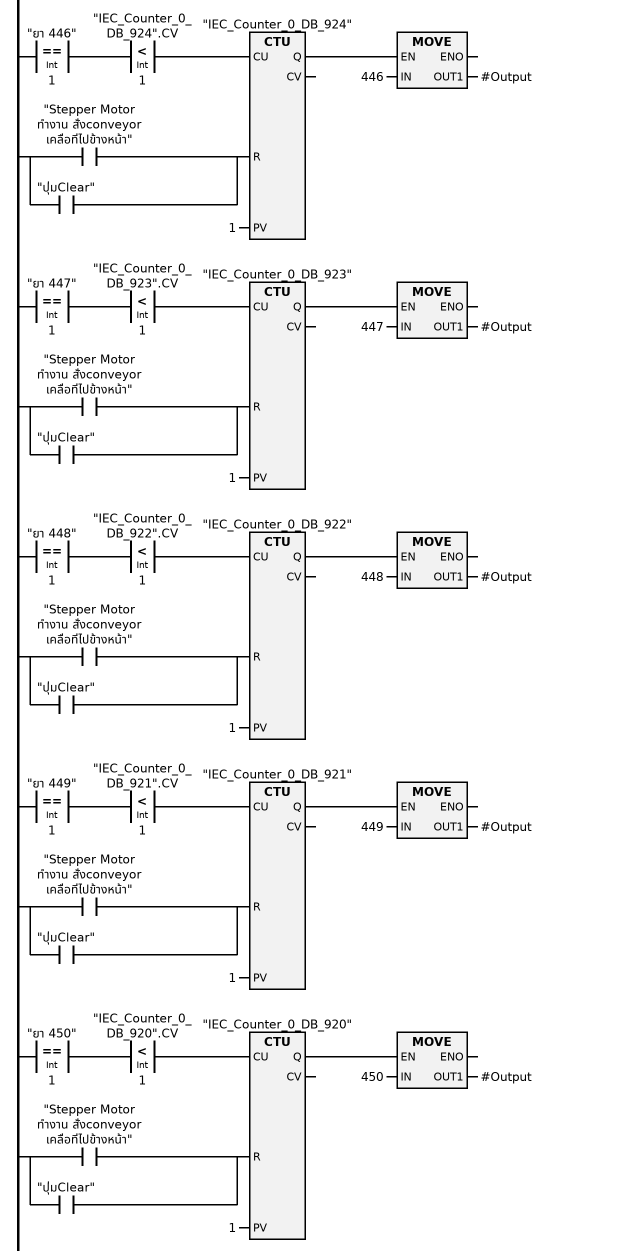
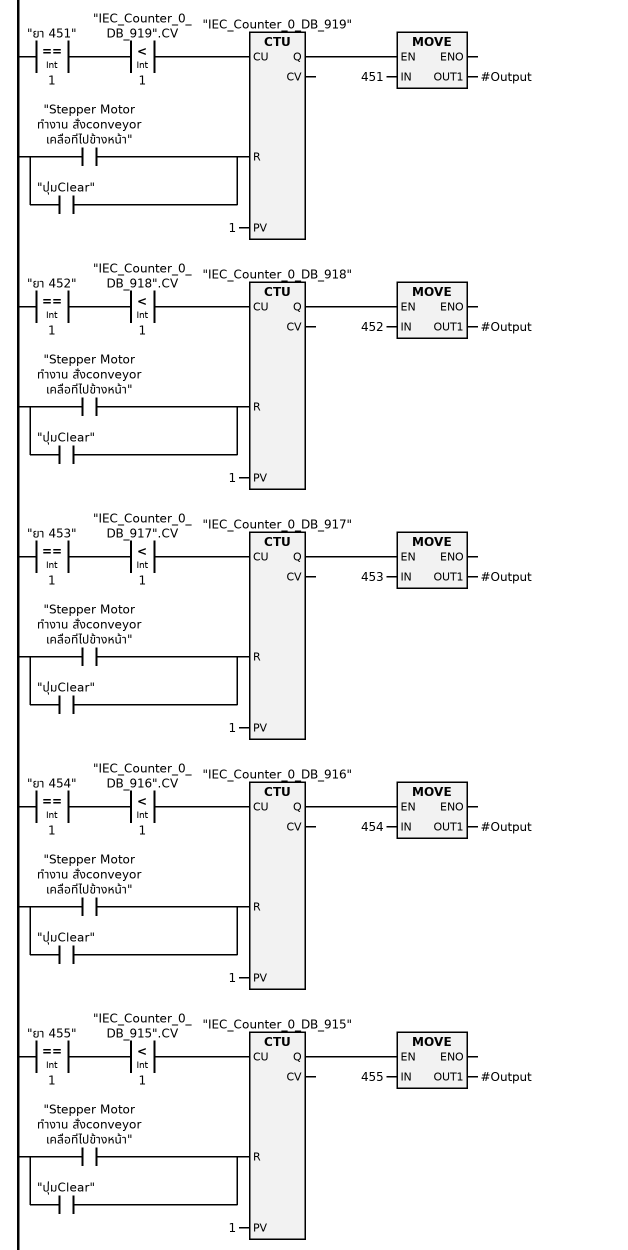
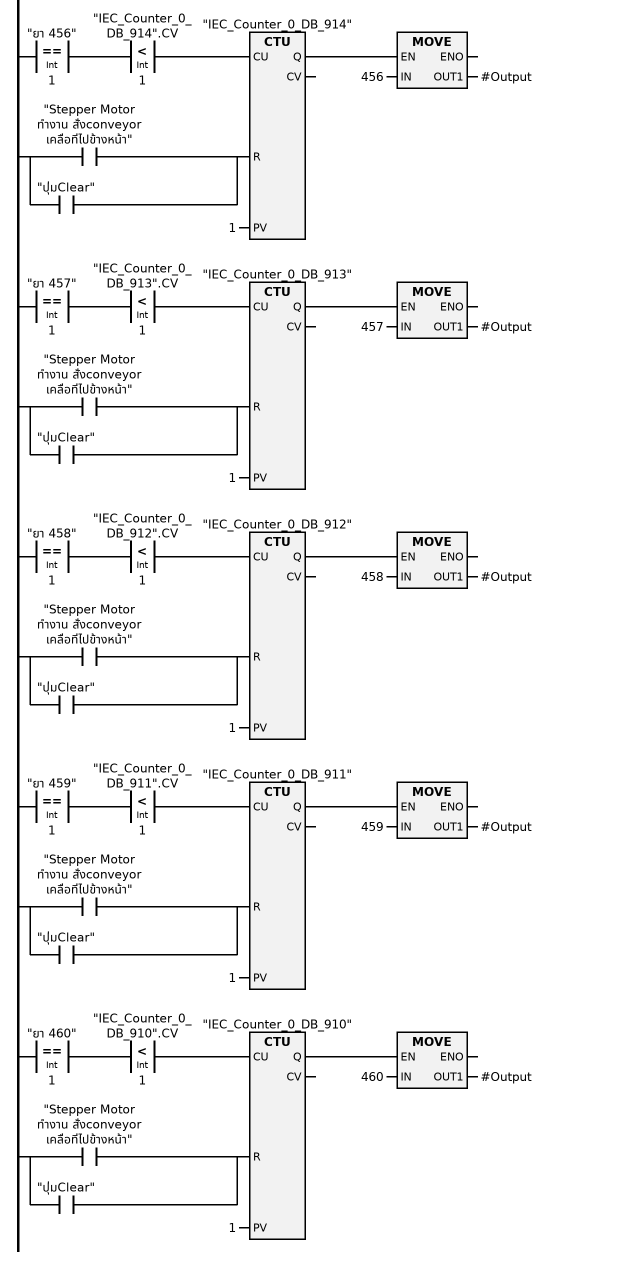
   "IEC_Counter_0_DB_929".CTU(CU := ("ยา 441" = 1) AND ("IEC_Counter_0_DB_929".CV < 1),
                           R := "Stepper Motor ทำงาน สั่งconveyor เคลื่อที่ไปข้างหน้า" OR "ปุ่มClear",
                           PV := 1);
   IF "IEC_Counter_0_DB_929".Q THEN #Output := 441; END_IF;
   "IEC_Counter_0_DB_928".CTU(CU := ("ยา 442" = 1) AND ("IEC_Counter_0_DB_928".CV < 1),
                           R := "Stepper Motor ทำงาน สั่งconveyor เคลื่อที่ไปข้างหน้า" OR "ปุ่มClear",
                           PV := 1);
   IF "IEC_Counter_0_DB_928".Q THEN #Output := 442; END_IF;
   "IEC_Counter_0_DB_927".CTU(CU := ("ยา 443" = 1) AND ("IEC_Counter_0_DB_927".CV < 1),
                           R := "Stepper Motor ทำงาน สั่งconveyor เคลื่อที่ไปข้างหน้า" OR "ปุ่มClear",
                           PV := 1);
   IF "IEC_Counter_0_DB_927".Q THEN #Output := 443; END_IF;
   "IEC_Counter_0_DB_926".CTU(CU := ("ยา 444" = 1) AND ("IEC_Counter_0_DB_926".CV < 1),
                           R := "Stepper Motor ทำงาน สั่งconveyor เคลื่อที่ไปข้างหน้า" OR "ปุ่มClear",
                           PV := 1);
   IF "IEC_Counter_0_DB_926".Q THEN #Output := 444; END_IF;
   "IEC_Counter_0_DB_925".CTU(CU := ("ยา 445" = 1) AND ("IEC_Counter_0_DB_925".CV < 1),
                           R := "Stepper Motor ทำงาน สั่งconveyor เคลื่อที่ไปข้างหน้า" OR "ปุ่มClear",
                           PV := 1);
   IF "IEC_Counter_0_DB_925".Q THEN #Output := 445; END_IF;
   "IEC_Counter_0_DB_924".CTU(CU := ("ยา 446" = 1) AND ("IEC_Counter_0_DB_924".CV < 1),
                           R := "Stepper Motor ทำงาน สั่งconveyor เคลื่อที่ไปข้างหน้า" OR "ปุ่มClear",
                           PV := 1);
   IF "IEC_Counter_0_DB_924".Q THEN #Output := 446; END_IF;
   "IEC_Counter_0_DB_923".CTU(CU := ("ยา 447" = 1) AND ("IEC_Counter_0_DB_923".CV < 1),
                           R := "Stepper Motor ทำงาน สั่งconveyor เคลื่อที่ไปข้างหน้า" OR "ปุ่มClear",
                           PV := 1);
   IF "IEC_Counter_0_DB_923".Q THEN #Output := 447; END_IF;
   "IEC_Counter_0_DB_922".CTU(CU := ("ยา 448" = 1) AND ("IEC_Counter_0_DB_922".CV < 1),
                           R := "Stepper Motor ทำงาน สั่งconveyor เคลื่อที่ไปข้างหน้า" OR "ปุ่มClear",
                           PV := 1);
   IF "IEC_Counter_0_DB_922".Q THEN #Output := 448; END_IF;
   "IEC_Counter_0_DB_921".CTU(CU := ("ยา 449" = 1) AND ("IEC_Counter_0_DB_921".CV < 1),
                           R := "Stepper Motor ทำงาน สั่งconveyor เคลื่อที่ไปข้างหน้า" OR "ปุ่มClear",
                           PV := 1);
   IF "IEC_Counter_0_DB_921".Q THEN #Output := 449; END_IF;
   "IEC_Counter_0_DB_920".CTU(CU := ("ยา 450" = 1) AND ("IEC_Counter_0_DB_920".CV < 1),
                           R := "Stepper Motor ทำงาน สั่งconveyor เคลื่อที่ไปข้างหน้า" OR "ปุ่มClear",
                           PV := 1);
   IF "IEC_Counter_0_DB_920".Q THEN #Output := 450; END_IF;
   "IEC_Counter_0_DB_919".CTU(CU := ("ยา 451" = 1) AND ("IEC_Counter_0_DB_919".CV < 1),
                           R := "Stepper Motor ทำงาน สั่งconveyor เคลื่อที่ไปข้างหน้า" OR "ปุ่มClear",
                           PV := 1);
   IF "IEC_Counter_0_DB_919".Q THEN #Output := 451; END_IF;
   "IEC_Counter_0_DB_918".CTU(CU := ("ยา 452" = 1) AND ("IEC_Counter_0_DB_918".CV < 1),
                           R := "Stepper Motor ทำงาน สั่งconveyor เคลื่อที่ไปข้างหน้า" OR "ปุ่มClear",
                           PV := 1);
   IF "IEC_Counter_0_DB_918".Q THEN #Output := 452; END_IF;
   "IEC_Counter_0_DB_917".CTU(CU := ("ยา 453" = 1) AND ("IEC_Counter_0_DB_917".CV < 1),
                           R := "Stepper Motor ทำงาน สั่งconveyor เคลื่อที่ไปข้างหน้า" OR "ปุ่มClear",
                           PV := 1);
   IF "IEC_Counter_0_DB_917".Q THEN #Output := 453; END_IF;
   "IEC_Counter_0_DB_916".CTU(CU := ("ยา 454" = 1) AND ("IEC_Counter_0_DB_916".CV < 1),
                           R := "Stepper Motor ทำงาน สั่งconveyor เคลื่อที่ไปข้างหน้า" OR "ปุ่มClear",
                           PV := 1);
   IF "IEC_Counter_0_DB_916".Q THEN #Output := 454; END_IF;
   "IEC_Counter_0_DB_915".CTU(CU := ("ยา 455" = 1) AND ("IEC_Counter_0_DB_915".CV < 1),
                           R := "Stepper Motor ทำงาน สั่งconveyor เคลื่อที่ไปข้างหน้า" OR "ปุ่มClear",
                           PV := 1);
   IF "IEC_Counter_0_DB_915".Q THEN #Output := 455; END_IF;
   "IEC_Counter_0_DB_914".CTU(CU := ("ยา 456" = 1) AND ("IEC_Counter_0_DB_914".CV < 1),
                           R := "Stepper Motor ทำงาน สั่งconveyor เคลื่อที่ไปข้างหน้า" OR "ปุ่มClear",
                           PV := 1);
   IF "IEC_Counter_0_DB_914".Q THEN #Output := 456; END_IF;
   "IEC_Counter_0_DB_913".CTU(CU := ("ยา 457" = 1) AND ("IEC_Counter_0_DB_913".CV < 1),
                           R := "Stepper Motor ทำงาน สั่งconveyor เคลื่อที่ไปข้างหน้า" OR "ปุ่มClear",
                           PV := 1);
   IF "IEC_Counter_0_DB_913".Q THEN #Output := 457; END_IF;
   "IEC_Counter_0_DB_912".CTU(CU := ("ยา 458" = 1) AND ("IEC_Counter_0_DB_912".CV < 1),
                           R := "Stepper Motor ทำงาน สั่งconveyor เคลื่อที่ไปข้างหน้า" OR "ปุ่มClear",
                           PV := 1);
   IF "IEC_Counter_0_DB_912".Q THEN #Output := 458; END_IF;
   "IEC_Counter_0_DB_911".CTU(CU := ("ยา 459" = 1) AND ("IEC_Counter_0_DB_911".CV < 1),
                           R := "Stepper Motor ทำงาน สั่งconveyor เคลื่อที่ไปข้างหน้า" OR "ปุ่มClear",
                           PV := 1);
   IF "IEC_Counter_0_DB_911".Q THEN #Output := 459; END_IF;
   "IEC_Counter_0_DB_910".CTU(CU := ("ยา 460" = 1) AND ("IEC_Counter_0_DB_910".CV < 1),
                           R := "Stepper Motor ทำงาน สั่งconveyor เคลื่อที่ไปข้างหน้า" OR "ปุ่มClear",
                           PV := 1);
   IF "IEC_Counter_0_DB_910".Q THEN #Output := 460; END_IF;
END_REGION

REGION Network 24
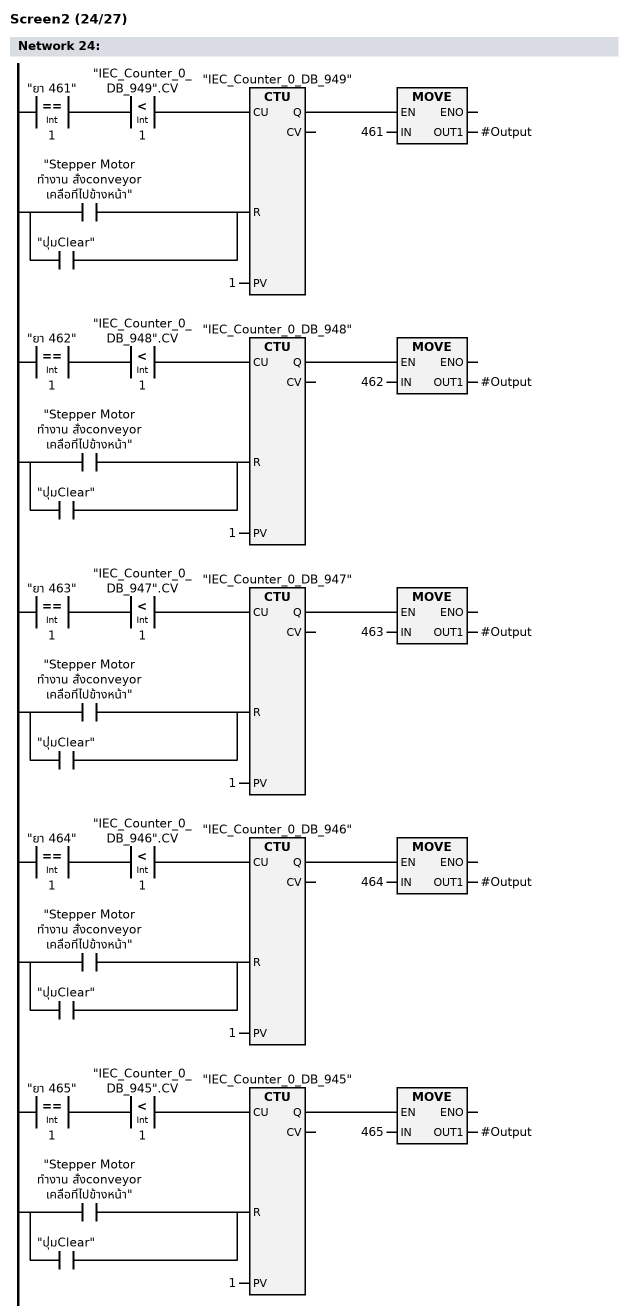
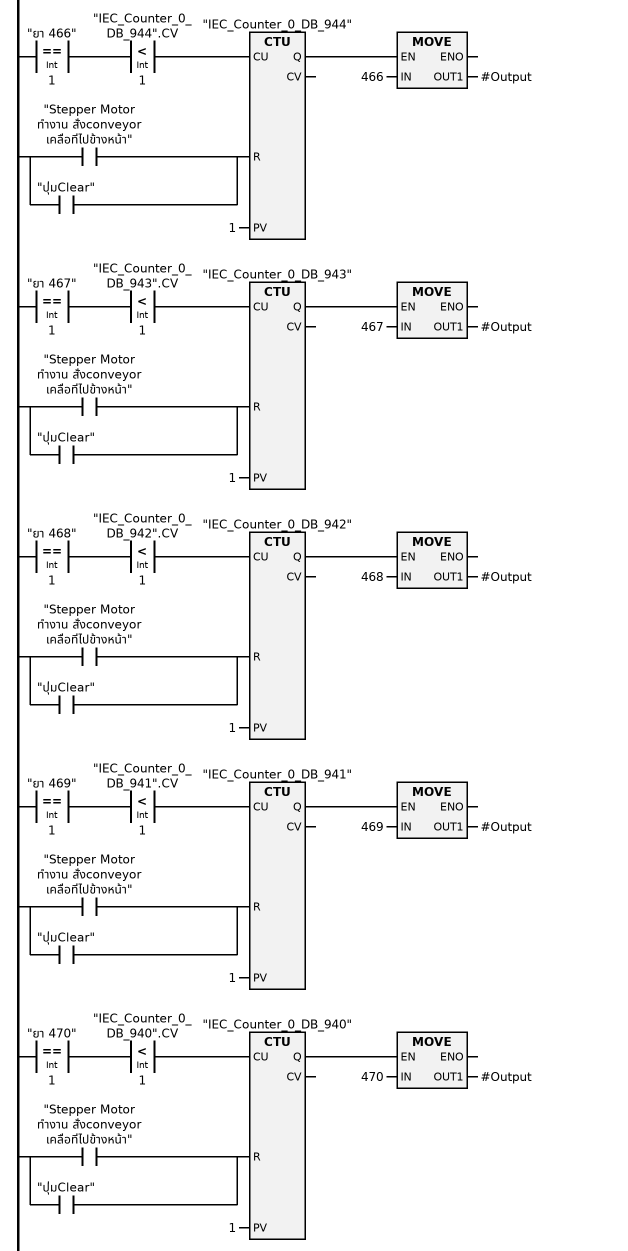
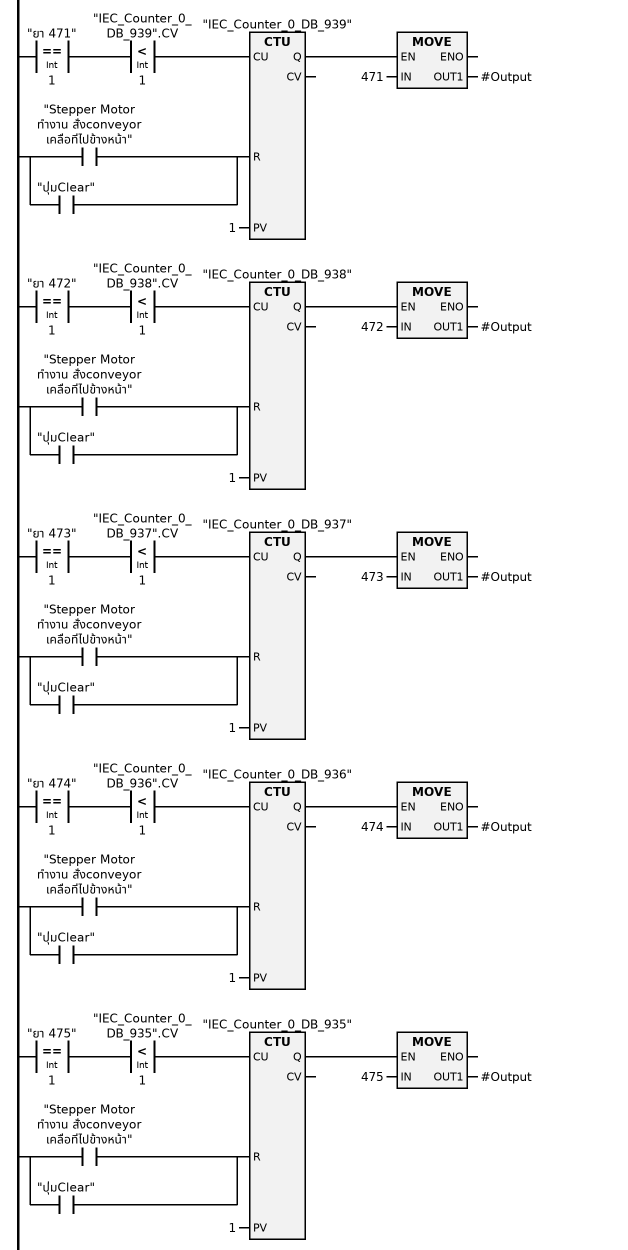
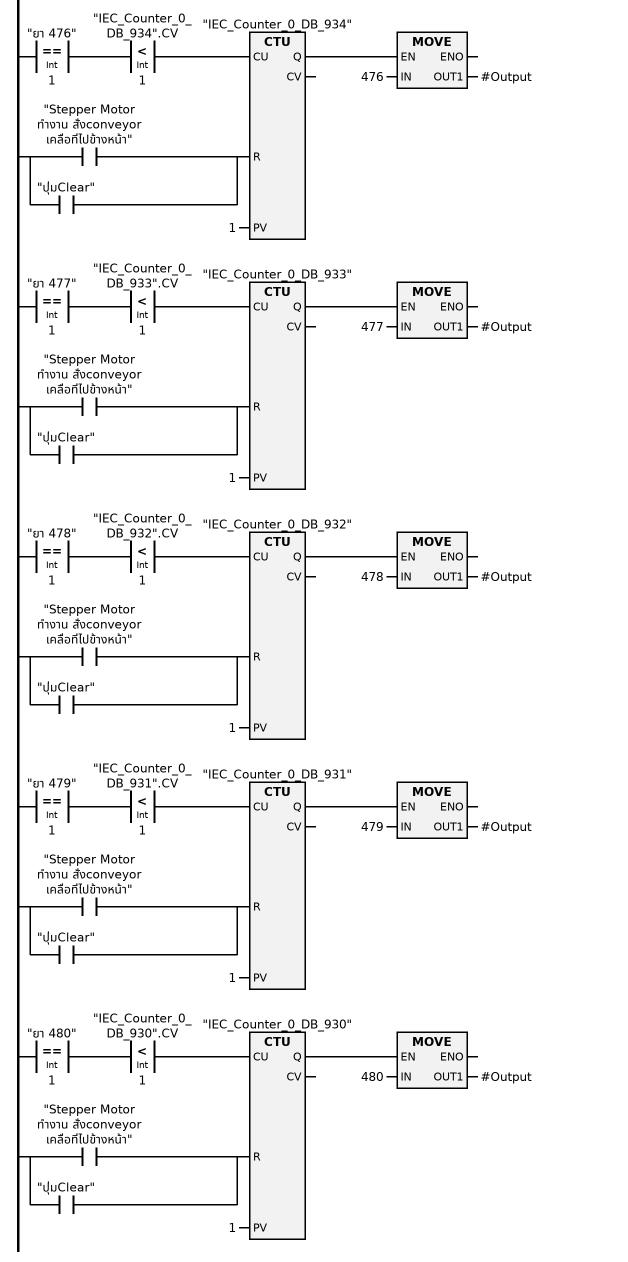
   "IEC_Counter_0_DB_949".CTU(CU := ("ยา 461" = 1) AND ("IEC_Counter_0_DB_949".CV < 1),
                           R := "Stepper Motor ทำงาน สั่งconveyor เคลื่อที่ไปข้างหน้า" OR "ปุ่มClear",
                           PV := 1);
   IF "IEC_Counter_0_DB_949".Q THEN #Output := 461; END_IF;
   "IEC_Counter_0_DB_948".CTU(CU := ("ยา 462" = 1) AND ("IEC_Counter_0_DB_948".CV < 1),
                           R := "Stepper Motor ทำงาน สั่งconveyor เคลื่อที่ไปข้างหน้า" OR "ปุ่มClear",
                           PV := 1);
   IF "IEC_Counter_0_DB_948".Q THEN #Output := 462; END_IF;
   "IEC_Counter_0_DB_947".CTU(CU := ("ยา 463" = 1) AND ("IEC_Counter_0_DB_947".CV < 1),
                           R := "Stepper Motor ทำงาน สั่งconveyor เคลื่อที่ไปข้างหน้า" OR "ปุ่มClear",
                           PV := 1);
   IF "IEC_Counter_0_DB_947".Q THEN #Output := 463; END_IF;
   "IEC_Counter_0_DB_946".CTU(CU := ("ยา 464" = 1) AND ("IEC_Counter_0_DB_946".CV < 1),
                           R := "Stepper Motor ทำงาน สั่งconveyor เคลื่อที่ไปข้างหน้า" OR "ปุ่มClear",
                           PV := 1);
   IF "IEC_Counter_0_DB_946".Q THEN #Output := 464; END_IF;
   "IEC_Counter_0_DB_945".CTU(CU := ("ยา 465" = 1) AND ("IEC_Counter_0_DB_945".CV < 1),
                           R := "Stepper Motor ทำงาน สั่งconveyor เคลื่อที่ไปข้างหน้า" OR "ปุ่มClear",
                           PV := 1);
   IF "IEC_Counter_0_DB_945".Q THEN #Output := 465; END_IF;
   "IEC_Counter_0_DB_944".CTU(CU := ("ยา 466" = 1) AND ("IEC_Counter_0_DB_944".CV < 1),
                           R := "Stepper Motor ทำงาน สั่งconveyor เคลื่อที่ไปข้างหน้า" OR "ปุ่มClear",
                           PV := 1);
   IF "IEC_Counter_0_DB_944".Q THEN #Output := 466; END_IF;
   "IEC_Counter_0_DB_943".CTU(CU := ("ยา 467" = 1) AND ("IEC_Counter_0_DB_943".CV < 1),
                           R := "Stepper Motor ทำงาน สั่งconveyor เคลื่อที่ไปข้างหน้า" OR "ปุ่มClear",
                           PV := 1);
   IF "IEC_Counter_0_DB_943".Q THEN #Output := 467; END_IF;
   "IEC_Counter_0_DB_942".CTU(CU := ("ยา 468" = 1) AND ("IEC_Counter_0_DB_942".CV < 1),
                           R := "Stepper Motor ทำงาน สั่งconveyor เคลื่อที่ไปข้างหน้า" OR "ปุ่มClear",
                           PV := 1);
   IF "IEC_Counter_0_DB_942".Q THEN #Output := 468; END_IF;
   "IEC_Counter_0_DB_941".CTU(CU := ("ยา 469" = 1) AND ("IEC_Counter_0_DB_941".CV < 1),
                           R := "Stepper Motor ทำงาน สั่งconveyor เคลื่อที่ไปข้างหน้า" OR "ปุ่มClear",
                           PV := 1);
   IF "IEC_Counter_0_DB_941".Q THEN #Output := 469; END_IF;
   "IEC_Counter_0_DB_940".CTU(CU := ("ยา 470" = 1) AND ("IEC_Counter_0_DB_940".CV < 1),
                           R := "Stepper Motor ทำงาน สั่งconveyor เคลื่อที่ไปข้างหน้า" OR "ปุ่มClear",
                           PV := 1);
   IF "IEC_Counter_0_DB_940".Q THEN #Output := 470; END_IF;
   "IEC_Counter_0_DB_939".CTU(CU := ("ยา 471" = 1) AND ("IEC_Counter_0_DB_939".CV < 1),
                           R := "Stepper Motor ทำงาน สั่งconveyor เคลื่อที่ไปข้างหน้า" OR "ปุ่มClear",
                           PV := 1);
   IF "IEC_Counter_0_DB_939".Q THEN #Output := 471; END_IF;
   "IEC_Counter_0_DB_938".CTU(CU := ("ยา 472" = 1) AND ("IEC_Counter_0_DB_938".CV < 1),
                           R := "Stepper Motor ทำงาน สั่งconveyor เคลื่อที่ไปข้างหน้า" OR "ปุ่มClear",
                           PV := 1);
   IF "IEC_Counter_0_DB_938".Q THEN #Output := 472; END_IF;
   "IEC_Counter_0_DB_937".CTU(CU := ("ยา 473" = 1) AND ("IEC_Counter_0_DB_937".CV < 1),
                           R := "Stepper Motor ทำงาน สั่งconveyor เคลื่อที่ไปข้างหน้า" OR "ปุ่มClear",
                           PV := 1);
   IF "IEC_Counter_0_DB_937".Q THEN #Output := 473; END_IF;
   "IEC_Counter_0_DB_936".CTU(CU := ("ยา 474" = 1) AND ("IEC_Counter_0_DB_936".CV < 1),
                           R := "Stepper Motor ทำงาน สั่งconveyor เคลื่อที่ไปข้างหน้า" OR "ปุ่มClear",
                           PV := 1);
   IF "IEC_Counter_0_DB_936".Q THEN #Output := 474; END_IF;
   "IEC_Counter_0_DB_935".CTU(CU := ("ยา 475" = 1) AND ("IEC_Counter_0_DB_935".CV < 1),
                           R := "Stepper Motor ทำงาน สั่งconveyor เคลื่อที่ไปข้างหน้า" OR "ปุ่มClear",
                           PV := 1);
   IF "IEC_Counter_0_DB_935".Q THEN #Output := 475; END_IF;
   "IEC_Counter_0_DB_934".CTU(CU := ("ยา 476" = 1) AND ("IEC_Counter_0_DB_934".CV < 1),
                           R := "Stepper Motor ทำงาน สั่งconveyor เคลื่อที่ไปข้างหน้า" OR "ปุ่มClear",
                           PV := 1);
   IF "IEC_Counter_0_DB_934".Q THEN #Output := 476; END_IF;
   "IEC_Counter_0_DB_933".CTU(CU := ("ยา 477" = 1) AND ("IEC_Counter_0_DB_933".CV < 1),
                           R := "Stepper Motor ทำงาน สั่งconveyor เคลื่อที่ไปข้างหน้า" OR "ปุ่มClear",
                           PV := 1);
   IF "IEC_Counter_0_DB_933".Q THEN #Output := 477; END_IF;
   "IEC_Counter_0_DB_932".CTU(CU := ("ยา 478" = 1) AND ("IEC_Counter_0_DB_932".CV < 1),
                           R := "Stepper Motor ทำงาน สั่งconveyor เคลื่อที่ไปข้างหน้า" OR "ปุ่มClear",
                           PV := 1);
   IF "IEC_Counter_0_DB_932".Q THEN #Output := 478; END_IF;
   "IEC_Counter_0_DB_931".CTU(CU := ("ยา 479" = 1) AND ("IEC_Counter_0_DB_931".CV < 1),
                           R := "Stepper Motor ทำงาน สั่งconveyor เคลื่อที่ไปข้างหน้า" OR "ปุ่มClear",
                           PV := 1);
   IF "IEC_Counter_0_DB_931".Q THEN #Output := 479; END_IF;
   "IEC_Counter_0_DB_930".CTU(CU := ("ยา 480" = 1) AND ("IEC_Counter_0_DB_930".CV < 1),
                           R := "Stepper Motor ทำงาน สั่งconveyor เคลื่อที่ไปข้างหน้า" OR "ปุ่มClear",
                           PV := 1);
   IF "IEC_Counter_0_DB_930".Q THEN #Output := 480; END_IF;
END_REGION

REGION Network 25
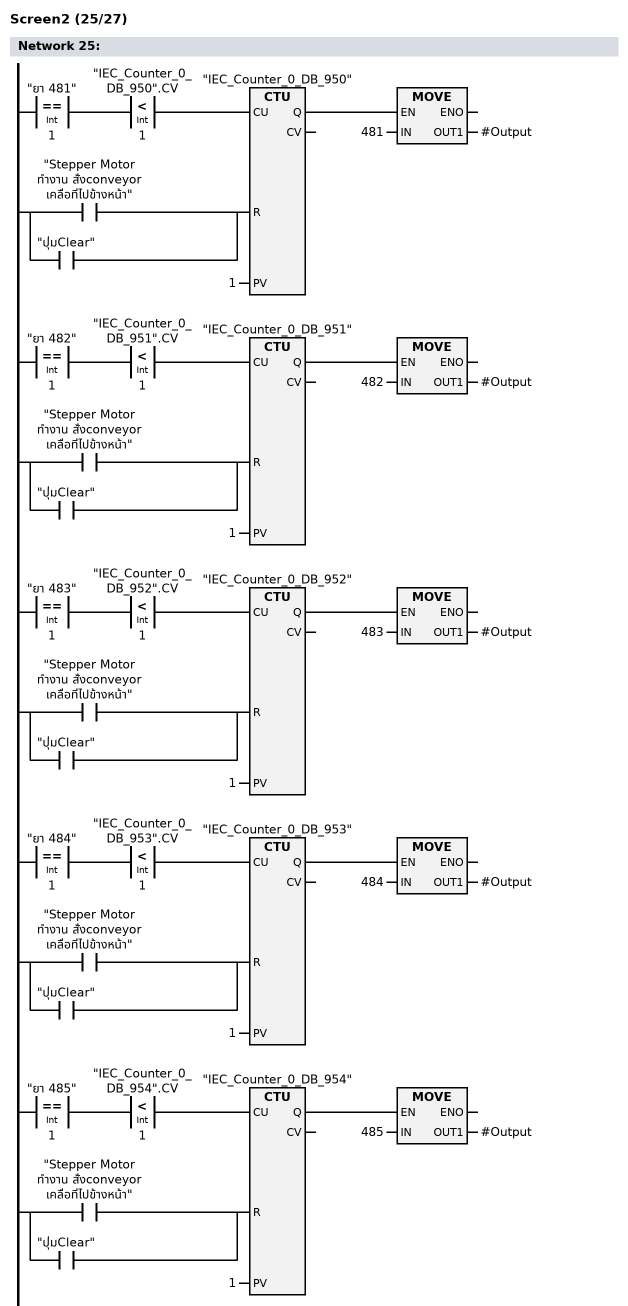
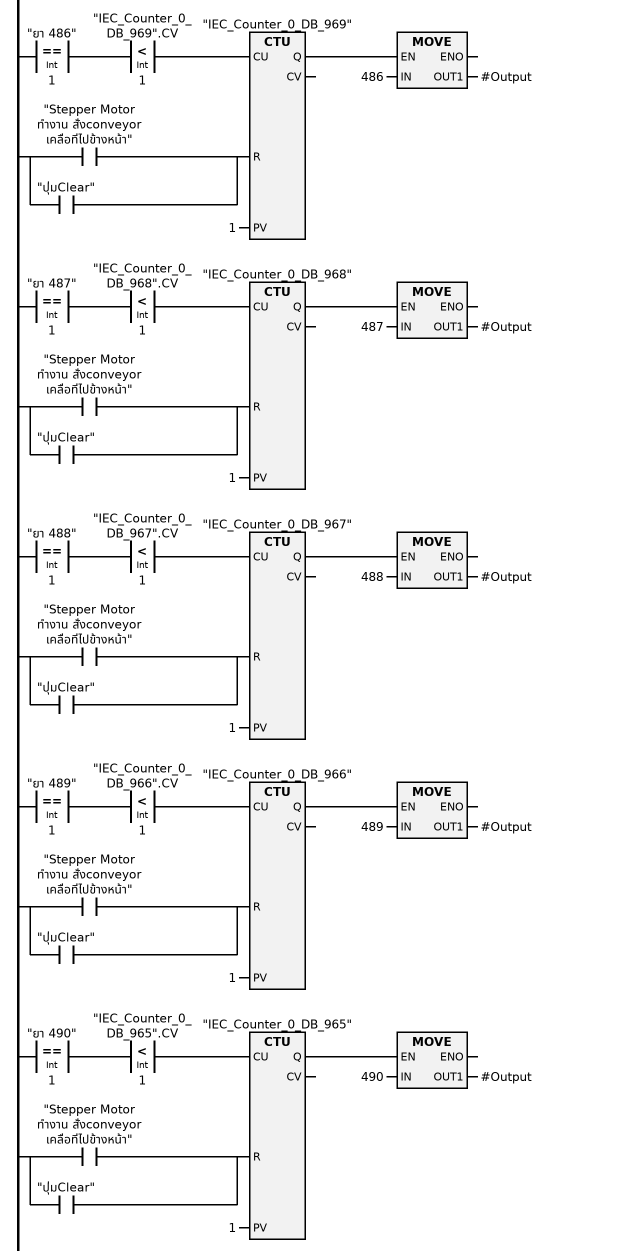
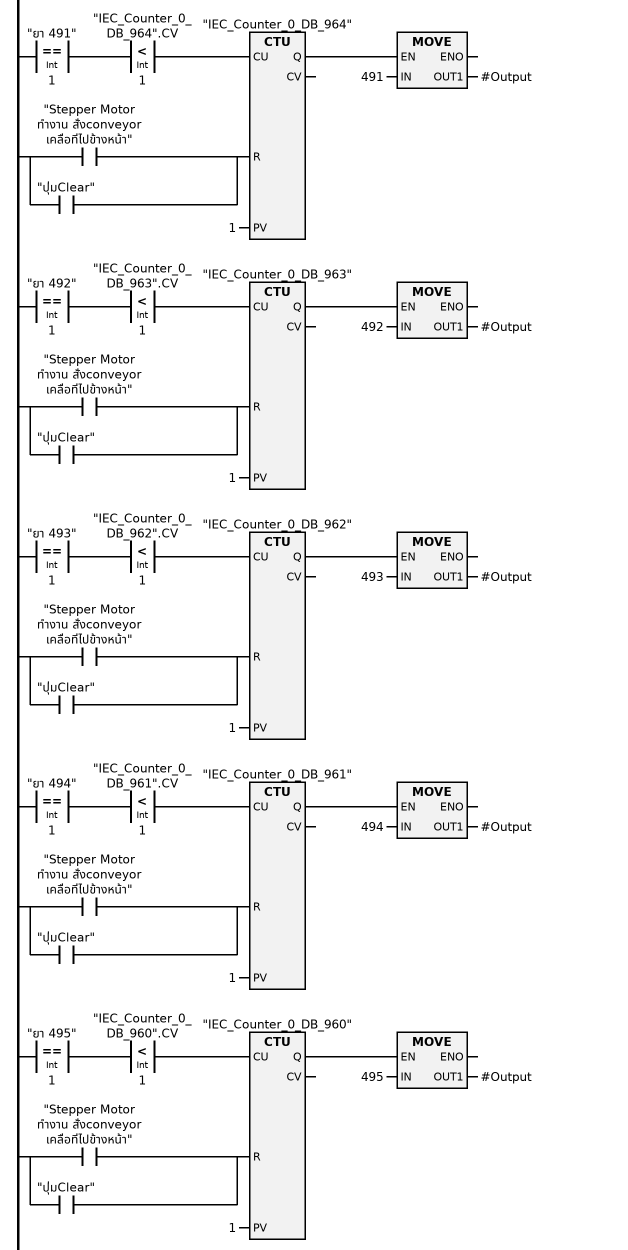
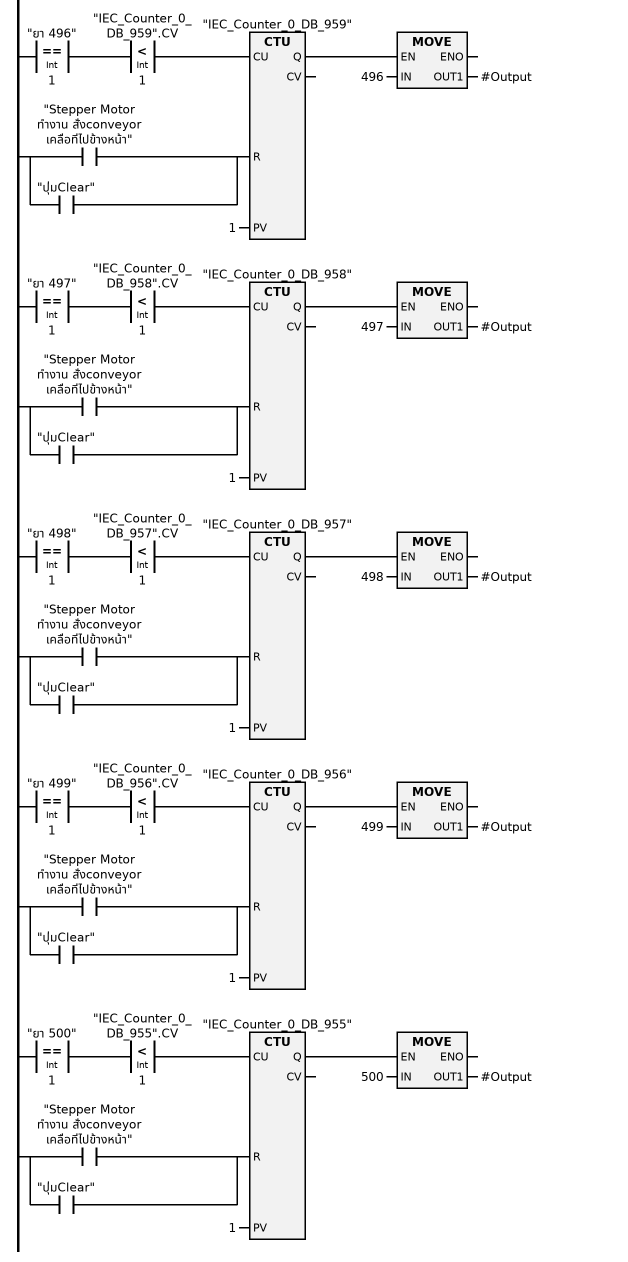
   "IEC_Counter_0_DB_950".CTU(CU := ("ยา 481" = 1) AND ("IEC_Counter_0_DB_950".CV < 1),
                           R := "Stepper Motor ทำงาน สั่งconveyor เคลื่อที่ไปข้างหน้า" OR "ปุ่มClear",
                           PV := 1);
   IF "IEC_Counter_0_DB_950".Q THEN #Output := 481; END_IF;
   "IEC_Counter_0_DB_951".CTU(CU := ("ยา 482" = 1) AND ("IEC_Counter_0_DB_951".CV < 1),
                           R := "Stepper Motor ทำงาน สั่งconveyor เคลื่อที่ไปข้างหน้า" OR "ปุ่มClear",
                           PV := 1);
   IF "IEC_Counter_0_DB_951".Q THEN #Output := 482; END_IF;
   "IEC_Counter_0_DB_952".CTU(CU := ("ยา 483" = 1) AND ("IEC_Counter_0_DB_952".CV < 1),
                           R := "Stepper Motor ทำงาน สั่งconveyor เคลื่อที่ไปข้างหน้า" OR "ปุ่มClear",
                           PV := 1);
   IF "IEC_Counter_0_DB_952".Q THEN #Output := 483; END_IF;
   "IEC_Counter_0_DB_953".CTU(CU := ("ยา 484" = 1) AND ("IEC_Counter_0_DB_953".CV < 1),
                           R := "Stepper Motor ทำงาน สั่งconveyor เคลื่อที่ไปข้างหน้า" OR "ปุ่มClear",
                           PV := 1);
   IF "IEC_Counter_0_DB_953".Q THEN #Output := 484; END_IF;
   "IEC_Counter_0_DB_954".CTU(CU := ("ยา 485" = 1) AND ("IEC_Counter_0_DB_954".CV < 1),
                           R := "Stepper Motor ทำงาน สั่งconveyor เคลื่อที่ไปข้างหน้า" OR "ปุ่มClear",
                           PV := 1);
   IF "IEC_Counter_0_DB_954".Q THEN #Output := 485; END_IF;
   "IEC_Counter_0_DB_969".CTU(CU := ("ยา 486" = 1) AND ("IEC_Counter_0_DB_969".CV < 1),
                           R := "Stepper Motor ทำงาน สั่งconveyor เคลื่อที่ไปข้างหน้า" OR "ปุ่มClear",
                           PV := 1);
   IF "IEC_Counter_0_DB_969".Q THEN #Output := 486; END_IF;
   "IEC_Counter_0_DB_968".CTU(CU := ("ยา 487" = 1) AND ("IEC_Counter_0_DB_968".CV < 1),
                           R := "Stepper Motor ทำงาน สั่งconveyor เคลื่อที่ไปข้างหน้า" OR "ปุ่มClear",
                           PV := 1);
   IF "IEC_Counter_0_DB_968".Q THEN #Output := 487; END_IF;
   "IEC_Counter_0_DB_967".CTU(CU := ("ยา 488" = 1) AND ("IEC_Counter_0_DB_967".CV < 1),
                           R := "Stepper Motor ทำงาน สั่งconveyor เคลื่อที่ไปข้างหน้า" OR "ปุ่มClear",
                           PV := 1);
   IF "IEC_Counter_0_DB_967".Q THEN #Output := 488; END_IF;
   "IEC_Counter_0_DB_966".CTU(CU := ("ยา 489" = 1) AND ("IEC_Counter_0_DB_966".CV < 1),
                           R := "Stepper Motor ทำงาน สั่งconveyor เคลื่อที่ไปข้างหน้า" OR "ปุ่มClear",
                           PV := 1);
   IF "IEC_Counter_0_DB_966".Q THEN #Output := 489; END_IF;
   "IEC_Counter_0_DB_965".CTU(CU := ("ยา 490" = 1) AND ("IEC_Counter_0_DB_965".CV < 1),
                           R := "Stepper Motor ทำงาน สั่งconveyor เคลื่อที่ไปข้างหน้า" OR "ปุ่มClear",
                           PV := 1);
   IF "IEC_Counter_0_DB_965".Q THEN #Output := 490; END_IF;
   "IEC_Counter_0_DB_964".CTU(CU := ("ยา 491" = 1) AND ("IEC_Counter_0_DB_964".CV < 1),
                           R := "Stepper Motor ทำงาน สั่งconveyor เคลื่อที่ไปข้างหน้า" OR "ปุ่มClear",
                           PV := 1);
   IF "IEC_Counter_0_DB_964".Q THEN #Output := 491; END_IF;
   "IEC_Counter_0_DB_963".CTU(CU := ("ยา 492" = 1) AND ("IEC_Counter_0_DB_963".CV < 1),
                           R := "Stepper Motor ทำงาน สั่งconveyor เคลื่อที่ไปข้างหน้า" OR "ปุ่มClear",
                           PV := 1);
   IF "IEC_Counter_0_DB_963".Q THEN #Output := 492; END_IF;
   "IEC_Counter_0_DB_962".CTU(CU := ("ยา 493" = 1) AND ("IEC_Counter_0_DB_962".CV < 1),
                           R := "Stepper Motor ทำงาน สั่งconveyor เคลื่อที่ไปข้างหน้า" OR "ปุ่มClear",
                           PV := 1);
   IF "IEC_Counter_0_DB_962".Q THEN #Output := 493; END_IF;
   "IEC_Counter_0_DB_961".CTU(CU := ("ยา 494" = 1) AND ("IEC_Counter_0_DB_961".CV < 1),
                           R := "Stepper Motor ทำงาน สั่งconveyor เคลื่อที่ไปข้างหน้า" OR "ปุ่มClear",
                           PV := 1);
   IF "IEC_Counter_0_DB_961".Q THEN #Output := 494; END_IF;
   "IEC_Counter_0_DB_960".CTU(CU := ("ยา 495" = 1) AND ("IEC_Counter_0_DB_960".CV < 1),
                           R := "Stepper Motor ทำงาน สั่งconveyor เคลื่อที่ไปข้างหน้า" OR "ปุ่มClear",
                           PV := 1);
   IF "IEC_Counter_0_DB_960".Q THEN #Output := 495; END_IF;
   "IEC_Counter_0_DB_959".CTU(CU := ("ยา 496" = 1) AND ("IEC_Counter_0_DB_959".CV < 1),
                           R := "Stepper Motor ทำงาน สั่งconveyor เคลื่อที่ไปข้างหน้า" OR "ปุ่มClear",
                           PV := 1);
   IF "IEC_Counter_0_DB_959".Q THEN #Output := 496; END_IF;
   "IEC_Counter_0_DB_958".CTU(CU := ("ยา 497" = 1) AND ("IEC_Counter_0_DB_958".CV < 1),
                           R := "Stepper Motor ทำงาน สั่งconveyor เคลื่อที่ไปข้างหน้า" OR "ปุ่มClear",
                           PV := 1);
   IF "IEC_Counter_0_DB_958".Q THEN #Output := 497; END_IF;
   "IEC_Counter_0_DB_957".CTU(CU := ("ยา 498" = 1) AND ("IEC_Counter_0_DB_957".CV < 1),
                           R := "Stepper Motor ทำงาน สั่งconveyor เคลื่อที่ไปข้างหน้า" OR "ปุ่มClear",
                           PV := 1);
   IF "IEC_Counter_0_DB_957".Q THEN #Output := 498; END_IF;
   "IEC_Counter_0_DB_956".CTU(CU := ("ยา 499" = 1) AND ("IEC_Counter_0_DB_956".CV < 1),
                           R := "Stepper Motor ทำงาน สั่งconveyor เคลื่อที่ไปข้างหน้า" OR "ปุ่มClear",
                           PV := 1);
   IF "IEC_Counter_0_DB_956".Q THEN #Output := 499; END_IF;
   "IEC_Counter_0_DB_955".CTU(CU := ("ยา 500" = 1) AND ("IEC_Counter_0_DB_955".CV < 1),
                           R := "Stepper Motor ทำงาน สั่งconveyor เคลื่อที่ไปข้างหน้า" OR "ปุ่มClear",
                           PV := 1);
   IF "IEC_Counter_0_DB_955".Q THEN #Output := 500; END_IF;
END_REGION

REGION Network 26
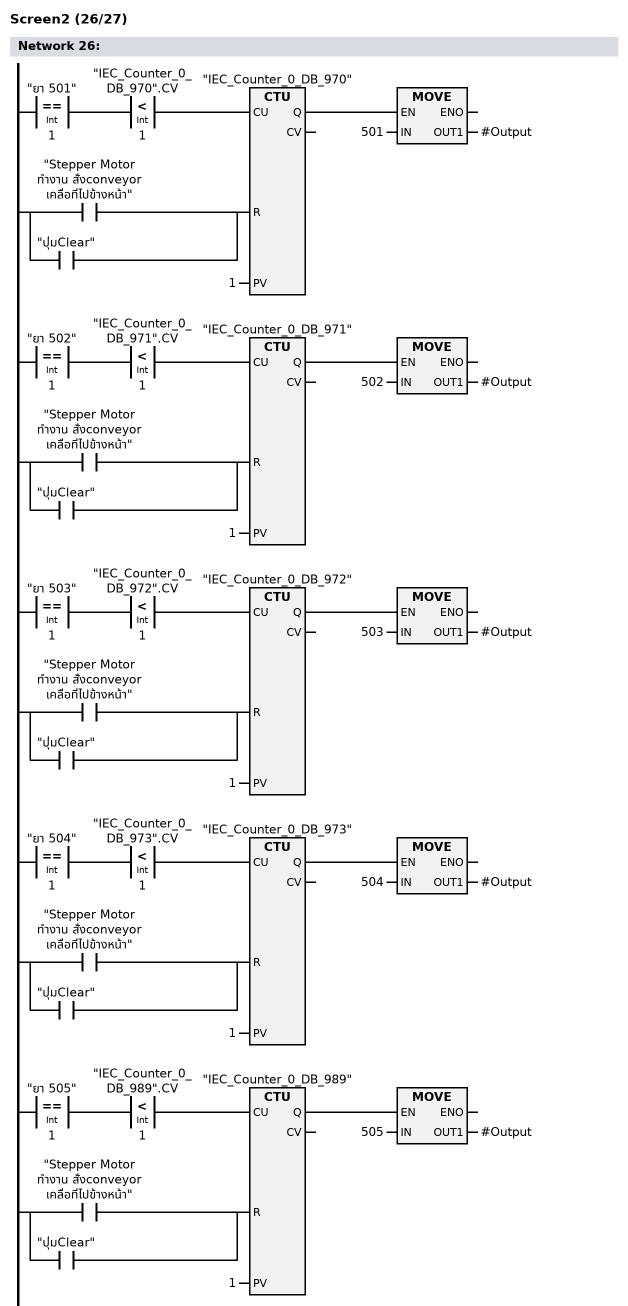
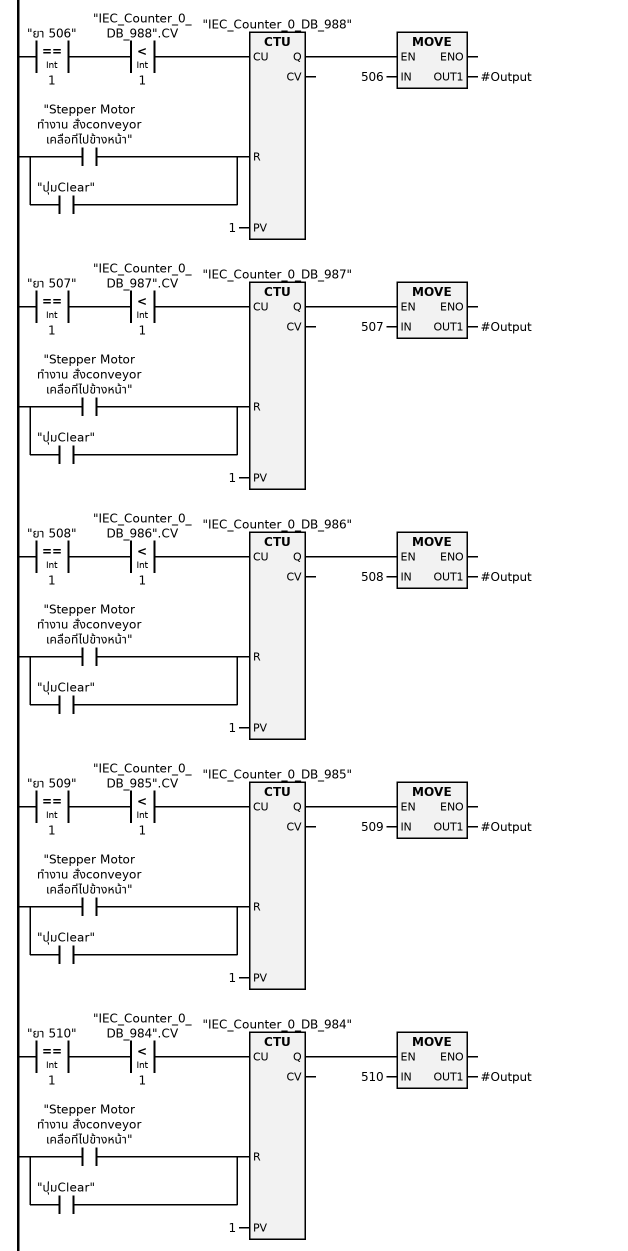
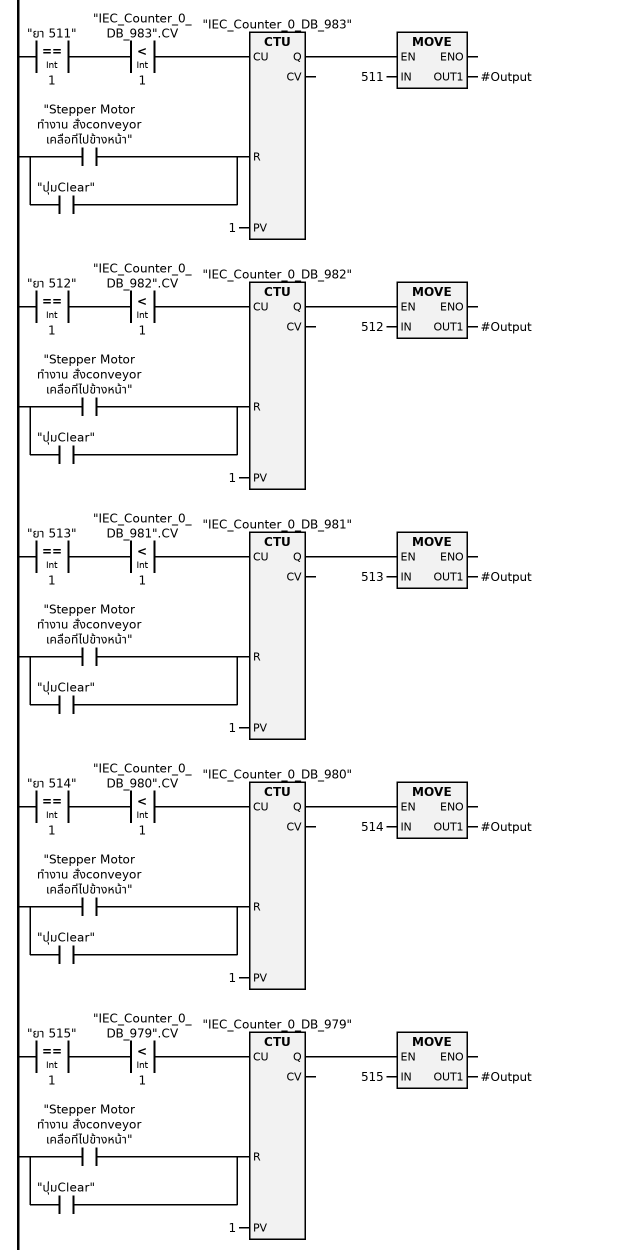
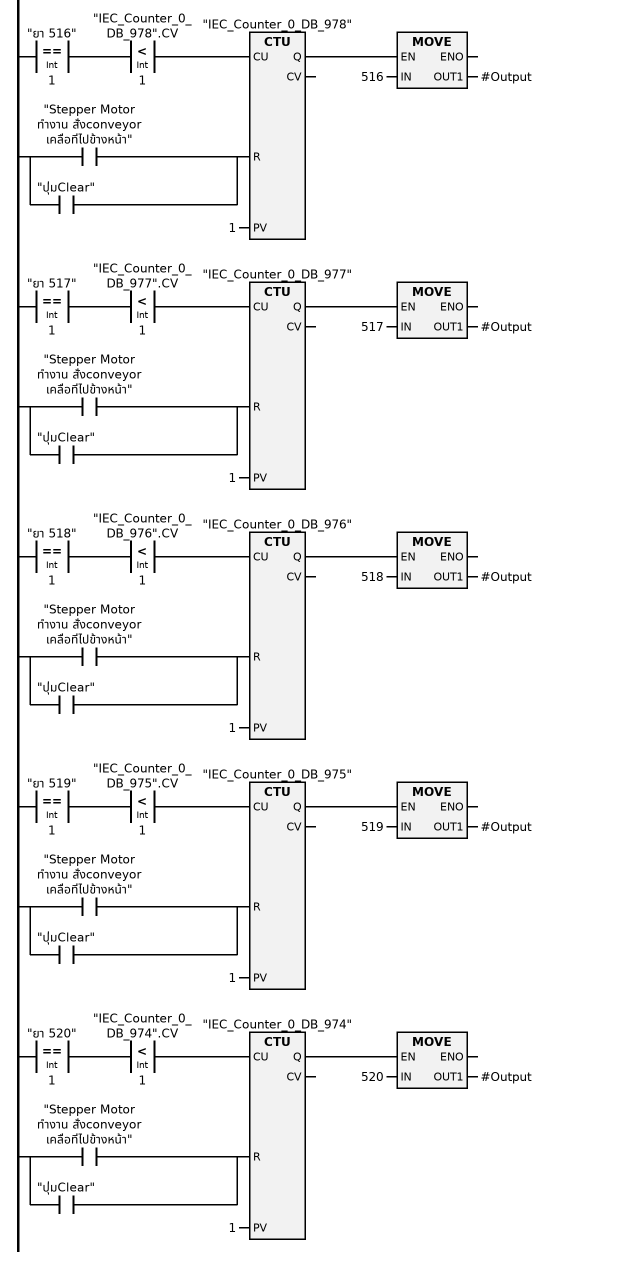
   "IEC_Counter_0_DB_970".CTU(CU := ("ยา 501" = 1) AND ("IEC_Counter_0_DB_970".CV < 1),
                           R := "Stepper Motor ทำงาน สั่งconveyor เคลื่อที่ไปข้างหน้า" OR "ปุ่มClear",
                           PV := 1);
   IF "IEC_Counter_0_DB_970".Q THEN #Output := 501; END_IF;
   "IEC_Counter_0_DB_971".CTU(CU := ("ยา 502" = 1) AND ("IEC_Counter_0_DB_971".CV < 1),
                           R := "Stepper Motor ทำงาน สั่งconveyor เคลื่อที่ไปข้างหน้า" OR "ปุ่มClear",
                           PV := 1);
   IF "IEC_Counter_0_DB_971".Q THEN #Output := 502; END_IF;
   "IEC_Counter_0_DB_972".CTU(CU := ("ยา 503" = 1) AND ("IEC_Counter_0_DB_972".CV < 1),
                           R := "Stepper Motor ทำงาน สั่งconveyor เคลื่อที่ไปข้างหน้า" OR "ปุ่มClear",
                           PV := 1);
   IF "IEC_Counter_0_DB_972".Q THEN #Output := 503; END_IF;
   "IEC_Counter_0_DB_973".CTU(CU := ("ยา 504" = 1) AND ("IEC_Counter_0_DB_973".CV < 1),
                           R := "Stepper Motor ทำงาน สั่งconveyor เคลื่อที่ไปข้างหน้า" OR "ปุ่มClear",
                           PV := 1);
   IF "IEC_Counter_0_DB_973".Q THEN #Output := 504; END_IF;
   "IEC_Counter_0_DB_989".CTU(CU := ("ยา 505" = 1) AND ("IEC_Counter_0_DB_989".CV < 1),
                           R := "Stepper Motor ทำงาน สั่งconveyor เคลื่อที่ไปข้างหน้า" OR "ปุ่มClear",
                           PV := 1);
   IF "IEC_Counter_0_DB_989".Q THEN #Output := 505; END_IF;
   "IEC_Counter_0_DB_988".CTU(CU := ("ยา 506" = 1) AND ("IEC_Counter_0_DB_988".CV < 1),
                           R := "Stepper Motor ทำงาน สั่งconveyor เคลื่อที่ไปข้างหน้า" OR "ปุ่มClear",
                           PV := 1);
   IF "IEC_Counter_0_DB_988".Q THEN #Output := 506; END_IF;
   "IEC_Counter_0_DB_987".CTU(CU := ("ยา 507" = 1) AND ("IEC_Counter_0_DB_987".CV < 1),
                           R := "Stepper Motor ทำงาน สั่งconveyor เคลื่อที่ไปข้างหน้า" OR "ปุ่มClear",
                           PV := 1);
   IF "IEC_Counter_0_DB_987".Q THEN #Output := 507; END_IF;
   "IEC_Counter_0_DB_986".CTU(CU := ("ยา 508" = 1) AND ("IEC_Counter_0_DB_986".CV < 1),
                           R := "Stepper Motor ทำงาน สั่งconveyor เคลื่อที่ไปข้างหน้า" OR "ปุ่มClear",
                           PV := 1);
   IF "IEC_Counter_0_DB_986".Q THEN #Output := 508; END_IF;
   "IEC_Counter_0_DB_985".CTU(CU := ("ยา 509" = 1) AND ("IEC_Counter_0_DB_985".CV < 1),
                           R := "Stepper Motor ทำงาน สั่งconveyor เคลื่อที่ไปข้างหน้า" OR "ปุ่มClear",
                           PV := 1);
   IF "IEC_Counter_0_DB_985".Q THEN #Output := 509; END_IF;
   "IEC_Counter_0_DB_984".CTU(CU := ("ยา 510" = 1) AND ("IEC_Counter_0_DB_984".CV < 1),
                           R := "Stepper Motor ทำงาน สั่งconveyor เคลื่อที่ไปข้างหน้า" OR "ปุ่มClear",
                           PV := 1);
   IF "IEC_Counter_0_DB_984".Q THEN #Output := 510; END_IF;
   "IEC_Counter_0_DB_983".CTU(CU := ("ยา 511" = 1) AND ("IEC_Counter_0_DB_983".CV < 1),
                           R := "Stepper Motor ทำงาน สั่งconveyor เคลื่อที่ไปข้างหน้า" OR "ปุ่มClear",
                           PV := 1);
   IF "IEC_Counter_0_DB_983".Q THEN #Output := 511; END_IF;
   "IEC_Counter_0_DB_982".CTU(CU := ("ยา 512" = 1) AND ("IEC_Counter_0_DB_982".CV < 1),
                           R := "Stepper Motor ทำงาน สั่งconveyor เคลื่อที่ไปข้างหน้า" OR "ปุ่มClear",
                           PV := 1);
   IF "IEC_Counter_0_DB_982".Q THEN #Output := 512; END_IF;
   "IEC_Counter_0_DB_981".CTU(CU := ("ยา 513" = 1) AND ("IEC_Counter_0_DB_981".CV < 1),
                           R := "Stepper Motor ทำงาน สั่งconveyor เคลื่อที่ไปข้างหน้า" OR "ปุ่มClear",
                           PV := 1);
   IF "IEC_Counter_0_DB_981".Q THEN #Output := 513; END_IF;
   "IEC_Counter_0_DB_980".CTU(CU := ("ยา 514" = 1) AND ("IEC_Counter_0_DB_980".CV < 1),
                           R := "Stepper Motor ทำงาน สั่งconveyor เคลื่อที่ไปข้างหน้า" OR "ปุ่มClear",
                           PV := 1);
   IF "IEC_Counter_0_DB_980".Q THEN #Output := 514; END_IF;
   "IEC_Counter_0_DB_979".CTU(CU := ("ยา 515" = 1) AND ("IEC_Counter_0_DB_979".CV < 1),
                           R := "Stepper Motor ทำงาน สั่งconveyor เคลื่อที่ไปข้างหน้า" OR "ปุ่มClear",
                           PV := 1);
   IF "IEC_Counter_0_DB_979".Q THEN #Output := 515; END_IF;
   "IEC_Counter_0_DB_978".CTU(CU := ("ยา 516" = 1) AND ("IEC_Counter_0_DB_978".CV < 1),
                           R := "Stepper Motor ทำงาน สั่งconveyor เคลื่อที่ไปข้างหน้า" OR "ปุ่มClear",
                           PV := 1);
   IF "IEC_Counter_0_DB_978".Q THEN #Output := 516; END_IF;
   "IEC_Counter_0_DB_977".CTU(CU := ("ยา 517" = 1) AND ("IEC_Counter_0_DB_977".CV < 1),
                           R := "Stepper Motor ทำงาน สั่งconveyor เคลื่อที่ไปข้างหน้า" OR "ปุ่มClear",
                           PV := 1);
   IF "IEC_Counter_0_DB_977".Q THEN #Output := 517; END_IF;
   "IEC_Counter_0_DB_976".CTU(CU := ("ยา 518" = 1) AND ("IEC_Counter_0_DB_976".CV < 1),
                           R := "Stepper Motor ทำงาน สั่งconveyor เคลื่อที่ไปข้างหน้า" OR "ปุ่มClear",
                           PV := 1);
   IF "IEC_Counter_0_DB_976".Q THEN #Output := 518; END_IF;
   "IEC_Counter_0_DB_975".CTU(CU := ("ยา 519" = 1) AND ("IEC_Counter_0_DB_975".CV < 1),
                           R := "Stepper Motor ทำงาน สั่งconveyor เคลื่อที่ไปข้างหน้า" OR "ปุ่มClear",
                           PV := 1);
   IF "IEC_Counter_0_DB_975".Q THEN #Output := 519; END_IF;
   "IEC_Counter_0_DB_974".CTU(CU := ("ยา 520" = 1) AND ("IEC_Counter_0_DB_974".CV < 1),
                           R := "Stepper Motor ทำงาน สั่งconveyor เคลื่อที่ไปข้างหน้า" OR "ปุ่มClear",
                           PV := 1);
   IF "IEC_Counter_0_DB_974".Q THEN #Output := 520; END_IF;
END_REGION

REGION Network 27
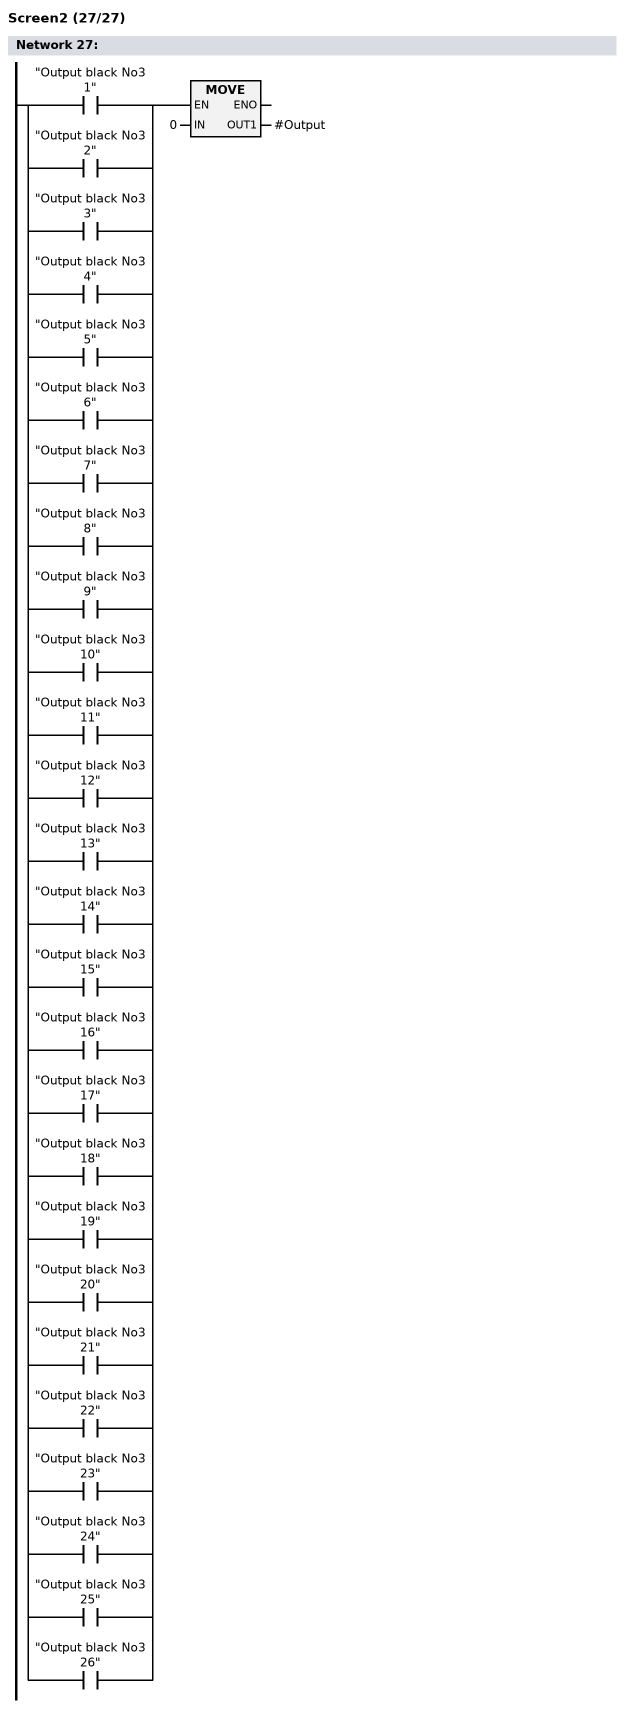
   RUNG wire#powerrail
      Contact( "Output black No3 1" )
      wire#w1
      Move(in := 0, out1 => #Output)
   END_RUNG
   RUNG wire#powerrail
      Contact( "Output black No3 2" )
   END_RUNG wire#w1
   RUNG wire#powerrail
      Contact( "Output black No3 3" )
   END_RUNG wire#w1
   RUNG wire#powerrail
      Contact( "Output black No3 4" )
   END_RUNG wire#w1
   RUNG wire#powerrail
      Contact( "Output black No3 5" )
   END_RUNG wire#w1
   RUNG wire#powerrail
      Contact( "Output black No3 6" )
   END_RUNG wire#w1
   RUNG wire#powerrail
      Contact( "Output black No3 7" )
   END_RUNG wire#w1
   RUNG wire#powerrail
      Contact( "Output black No3 8" )
   END_RUNG wire#w1
   RUNG wire#powerrail
      Contact( "Output black No3 9" )
   END_RUNG wire#w1
   RUNG wire#powerrail
      Contact( "Output black No3 10" )
   END_RUNG wire#w1
   RUNG wire#powerrail
      Contact( "Output black No3 11" )
   END_RUNG wire#w1
   RUNG wire#powerrail
      Contact( "Output black No3 12" )
   END_RUNG wire#w1
   RUNG wire#powerrail
      Contact( "Output black No3 13" )
   END_RUNG wire#w1
   RUNG wire#powerrail
      Contact( "Output black No3 14" )
   END_RUNG wire#w1
   RUNG wire#powerrail
      Contact( "Output black No3 15" )
   END_RUNG wire#w1
   RUNG wire#powerrail
      Contact( "Output black No3 16" )
   END_RUNG wire#w1
   RUNG wire#powerrail
      Contact( "Output black No3 17" )
   END_RUNG wire#w1
   RUNG wire#powerrail
      Contact( "Output black No3 18" )
   END_RUNG wire#w1
   RUNG wire#powerrail
      Contact( "Output black No3 19" )
   END_RUNG wire#w1
   RUNG wire#powerrail
      Contact( "Output black No3 20" )
   END_RUNG wire#w1
   RUNG wire#powerrail
      Contact( "Output black No3 21" )
   END_RUNG wire#w1
   RUNG wire#powerrail
      Contact( "Output black No3 22" )
   END_RUNG wire#w1
   RUNG wire#powerrail
      Contact( "Output black No3 23" )
   END_RUNG wire#w1
   RUNG wire#powerrail
      Contact( "Output black No3 24" )
   END_RUNG wire#w1
   RUNG wire#powerrail
      Contact( "Output black No3 25" )
   END_RUNG wire#w1
   RUNG wire#powerrail
      Contact( "Output black No3 26" )
   END_RUNG wire#w1
   // the same network as SCL:
   IF "Output black No3 1" OR "Output black No3 2" OR "Output black No3 3" OR "Output black No3 4" OR "Output black No3 5" OR "Output black No3 6" OR "Output black No3 7" OR "Output black No3 8" OR "Output black No3 9" OR "Output black No3 10" OR "Output black No3 11" OR "Output black No3 12" OR "Output black No3 13" OR "Output black No3 14" OR "Output black No3 15" OR "Output black No3 16" OR "Output black No3 17" OR "Output black No3 18" OR "Output black No3 19" OR "Output black No3 20" OR "Output black No3 21" OR "Output black No3 22" OR "Output black No3 23" OR "Output black No3 24" OR "Output black No3 25" OR "Output black No3 26" THEN
       #Output := 0;
   END_IF;
END_REGION
END_FUNCTION

FUNCTION "Screen3 Data เบิกจ่าย / จัดเก็บ" : Void   // FC15, LAD
{ S7_Optimized_Access := 'TRUE' }
VERSION : 0.1
   VAR_OUTPUT
      Output : Word;
      Output1 : Word;
      Output2 : Word;
      Output3 : Word;
   END_VAR
BEGIN

REGION Network 1: เบิกจ่าย
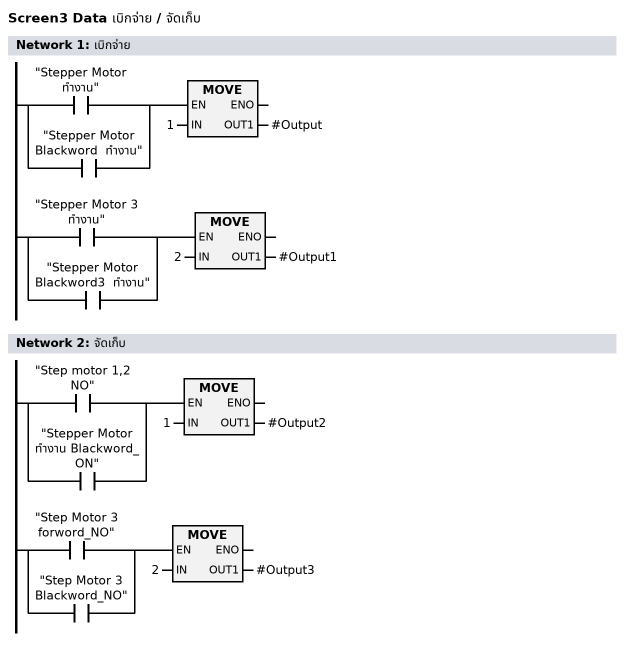
   RUNG wire#powerrail
      Contact( "Stepper Motor  ทำงาน" )
      wire#w1
      Move(in := 1, out1 => #Output)
   END_RUNG
   RUNG wire#powerrail
      Contact( "Stepper Motor Blackword  ทำงาน" )
   END_RUNG wire#w1
   RUNG wire#powerrail
      Contact( "Stepper Motor 3 ทำงาน" )
      wire#w2
      Move(in := 2, out1 => #Output1)
   END_RUNG
   RUNG wire#powerrail
      Contact( "Stepper Motor Blackword3  ทำงาน" )
   END_RUNG wire#w2
   // the same network as SCL:
   IF "Stepper Motor  ทำงาน" OR "Stepper Motor Blackword  ทำงาน" THEN #Output := 1; END_IF;
   IF "Stepper Motor 3 ทำงาน" OR "Stepper Motor Blackword3  ทำงาน" THEN #Output1 := 2; END_IF;
END_REGION

REGION Network 2: จัดเก็บ
   RUNG wire#powerrail
      Contact( "Step motor 1,2 NO" )
      wire#w1
      Move(in := 1, out1 => #Output2)
   END_RUNG
   RUNG wire#powerrail
      Contact( "Stepper Motor  ทำงาน Blackword_ON" )
   END_RUNG wire#w1
   RUNG wire#powerrail
      Contact( "Step Motor 3 forword_NO" )
      wire#w2
      Move(in := 2, out1 => #Output3)
   END_RUNG
   RUNG wire#powerrail
      Contact( "Step Motor 3 Blackword_NO" )
   END_RUNG wire#w2
   // the same network as SCL:
   IF "Step motor 1,2 NO" OR "Stepper Motor  ทำงาน Blackword_ON" THEN #Output2 := 1; END_IF;
   IF "Step Motor 3 forword_NO" OR "Step Motor 3 Blackword_NO" THEN #Output3 := 2; END_IF;
END_REGION
END_FUNCTION

FUNCTION "output Reset ชื่อยา" : Void   // FC16, LAD
{ S7_Optimized_Access := 'TRUE' }
VERSION : 0.1
BEGIN

REGION Network 1
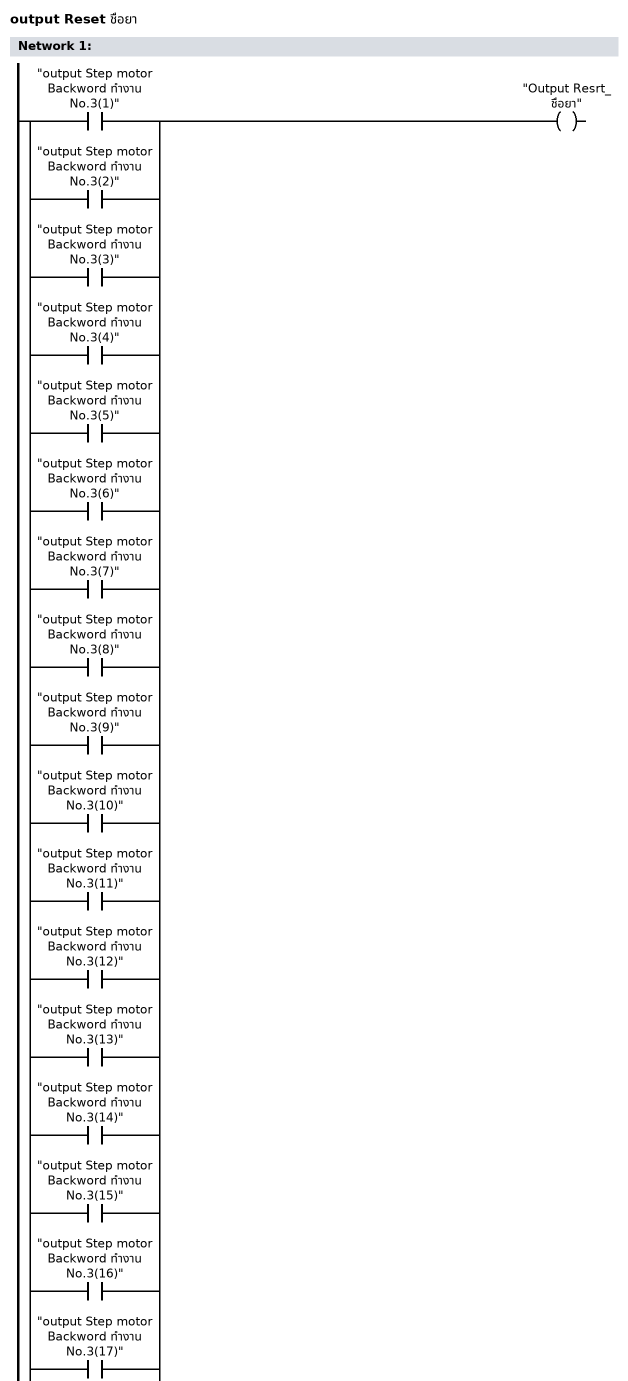
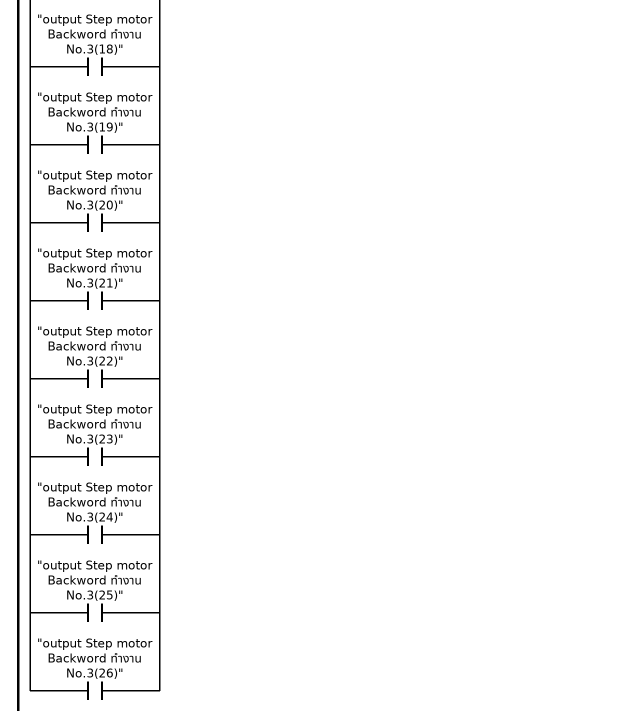
   RUNG wire#powerrail
      Contact( "output Step motor  Backword ทำงาน No.3(1)" )
      wire#w1
      Coil( "Output Resrt_ชื่อยา" )
   END_RUNG
   RUNG wire#powerrail
      Contact( "output Step motor  Backword ทำงาน No.3(2)" )
   END_RUNG wire#w1
   RUNG wire#powerrail
      Contact( "output Step motor  Backword ทำงาน No.3(3)" )
   END_RUNG wire#w1
   RUNG wire#powerrail
      Contact( "output Step motor  Backword ทำงาน No.3(4)" )
   END_RUNG wire#w1
   RUNG wire#powerrail
      Contact( "output Step motor  Backword ทำงาน No.3(5)" )
   END_RUNG wire#w1
   RUNG wire#powerrail
      Contact( "output Step motor  Backword ทำงาน No.3(6)" )
   END_RUNG wire#w1
   RUNG wire#powerrail
      Contact( "output Step motor  Backword ทำงาน No.3(7)" )
   END_RUNG wire#w1
   RUNG wire#powerrail
      Contact( "output Step motor  Backword ทำงาน No.3(8)" )
   END_RUNG wire#w1
   RUNG wire#powerrail
      Contact( "output Step motor  Backword ทำงาน No.3(9)" )
   END_RUNG wire#w1
   RUNG wire#powerrail
      Contact( "output Step motor  Backword ทำงาน No.3(10)" )
   END_RUNG wire#w1
   RUNG wire#powerrail
      Contact( "output Step motor  Backword ทำงาน No.3(11)" )
   END_RUNG wire#w1
   RUNG wire#powerrail
      Contact( "output Step motor  Backword ทำงาน No.3(12)" )
   END_RUNG wire#w1
   RUNG wire#powerrail
      Contact( "output Step motor  Backword ทำงาน No.3(13)" )
   END_RUNG wire#w1
   RUNG wire#powerrail
      Contact( "output Step motor  Backword ทำงาน No.3(14)" )
   END_RUNG wire#w1
   RUNG wire#powerrail
      Contact( "output Step motor  Backword ทำงาน No.3(15)" )
   END_RUNG wire#w1
   RUNG wire#powerrail
      Contact( "output Step motor  Backword ทำงาน No.3(16)" )
   END_RUNG wire#w1
   RUNG wire#powerrail
      Contact( "output Step motor  Backword ทำงาน No.3(17)" )
   END_RUNG wire#w1
   RUNG wire#powerrail
      Contact( "output Step motor  Backword ทำงาน No.3(18)" )
   END_RUNG wire#w1
   RUNG wire#powerrail
      Contact( "output Step motor  Backword ทำงาน No.3(19)" )
   END_RUNG wire#w1
   RUNG wire#powerrail
      Contact( "output Step motor  Backword ทำงาน No.3(20)" )
   END_RUNG wire#w1
   RUNG wire#powerrail
      Contact( "output Step motor  Backword ทำงาน No.3(21)" )
   END_RUNG wire#w1
   RUNG wire#powerrail
      Contact( "output Step motor  Backword ทำงาน No.3(22)" )
   END_RUNG wire#w1
   RUNG wire#powerrail
      Contact( "output Step motor  Backword ทำงาน No.3(23)" )
   END_RUNG wire#w1
   RUNG wire#powerrail
      Contact( "output Step motor  Backword ทำงาน No.3(24)" )
   END_RUNG wire#w1
   RUNG wire#powerrail
      Contact( "output Step motor  Backword ทำงาน No.3(25)" )
   END_RUNG wire#w1
   RUNG wire#powerrail
      Contact( "output Step motor  Backword ทำงาน No.3(26)" )
   END_RUNG wire#w1
   // the same network as SCL:
   "Output Resrt_ชื่อยา" := "output Step motor  Backword ทำงาน No.3(1)" OR "output Step motor  Backword ทำงาน No.3(2)" OR "output Step motor  Backword ทำงาน No.3(3)" OR "output Step motor  Backword ทำงาน No.3(4)" OR "output Step motor  Backword ทำงาน No.3(5)" OR "output Step motor  Backword ทำงาน No.3(6)" OR "output Step motor  Backword ทำงาน No.3(7)" OR "output Step motor  Backword ทำงาน No.3(8)" OR "output Step motor  Backword ทำงาน No.3(9)" OR "output Step motor  Backword ทำงาน No.3(10)" OR "output Step motor  Backword ทำงาน No.3(11)" OR "output Step motor  Backword ทำงาน No.3(12)" OR "output Step motor  Backword ทำงาน No.3(13)" OR "output Step motor  Backword ทำงาน No.3(14)" OR "output Step motor  Backword ทำงาน No.3(15)" OR "output Step motor  Backword ทำงาน No.3(16)" OR "output Step motor  Backword ทำงาน No.3(17)" OR "output Step motor  Backword ทำงาน No.3(18)" OR "output Step motor  Backword ทำงาน No.3(19)" OR "output Step motor  Backword ทำงาน No.3(20)" OR "output Step motor  Backword ทำงาน No.3(21)" OR "output Step motor  Backword ทำงาน No.3(22)" OR "output Step motor  Backword ทำงาน No.3(23)" OR "output Step motor  Backword ทำงาน No.3(24)" OR "output Step motor  Backword ทำงาน No.3(25)" OR "output Step motor  Backword ทำงาน No.3(26)";
END_REGION
END_FUNCTION

FUNCTION "Screen4 Status" : Void   // FC18, LAD
{ S7_Optimized_Access := 'TRUE' }
VERSION : 0.1
BEGIN

REGION Network 1: จัดเก็บ
   // รับคำสั่งจัดเก็บยา
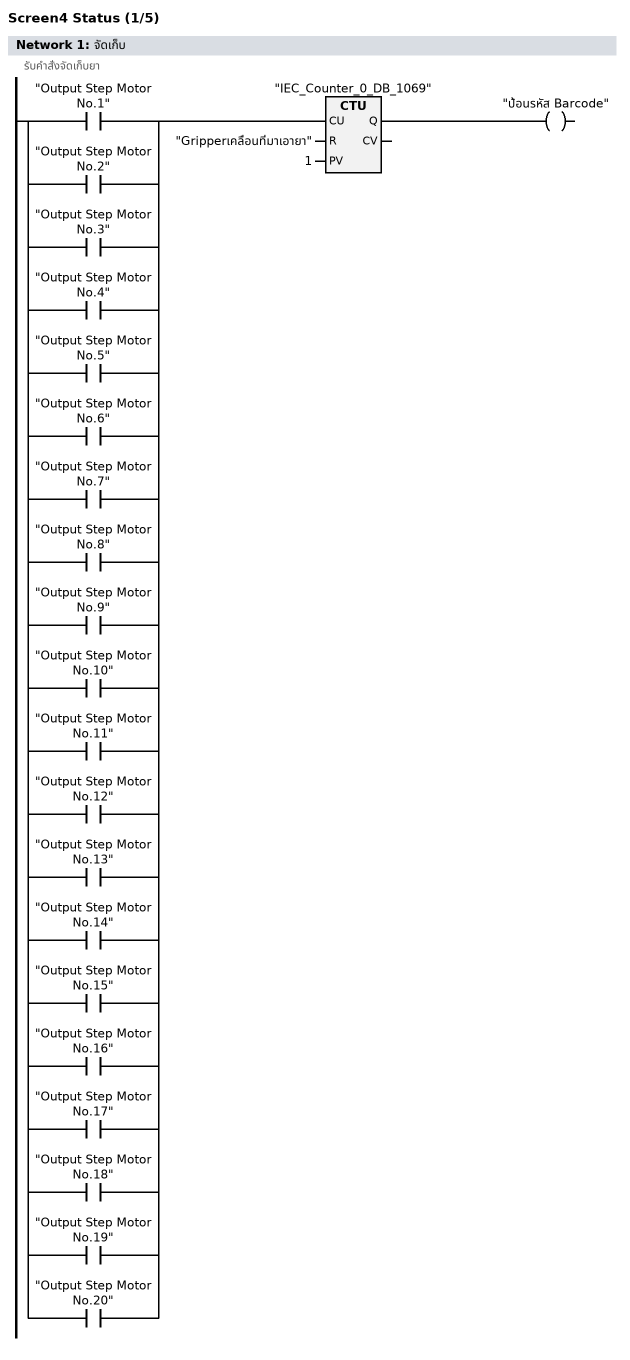
   "IEC_Counter_0_DB_1069".CTU(CU := "Output Step Motor No.1" OR "Output Step Motor No.2" OR "Output Step Motor No.3" OR "Output Step Motor No.4" OR "Output Step Motor No.5" OR "Output Step Motor No.6" OR "Output Step Motor No.7" OR "Output Step Motor No.8" OR "Output Step Motor No.9" OR "Output Step Motor No.10" OR "Output Step Motor No.11" OR "Output Step Motor No.12" OR "Output Step Motor No.13" OR "Output Step Motor No.14" OR "Output Step Motor No.15" OR "Output Step Motor No.16" OR "Output Step Motor No.17" OR "Output Step Motor No.18" OR "Output Step Motor No.19" OR "Output Step Motor No.20",
                           R := "Gripperเคลื่อนที่มาเอายา",
                           PV := 1);
   "ป้อนรหัส Barcode" := "IEC_Counter_0_DB_1069".Q;
END_REGION

REGION Network 2: จัดเก็บ
   // Gripperเคลื่อนที่
   //  มารับยา
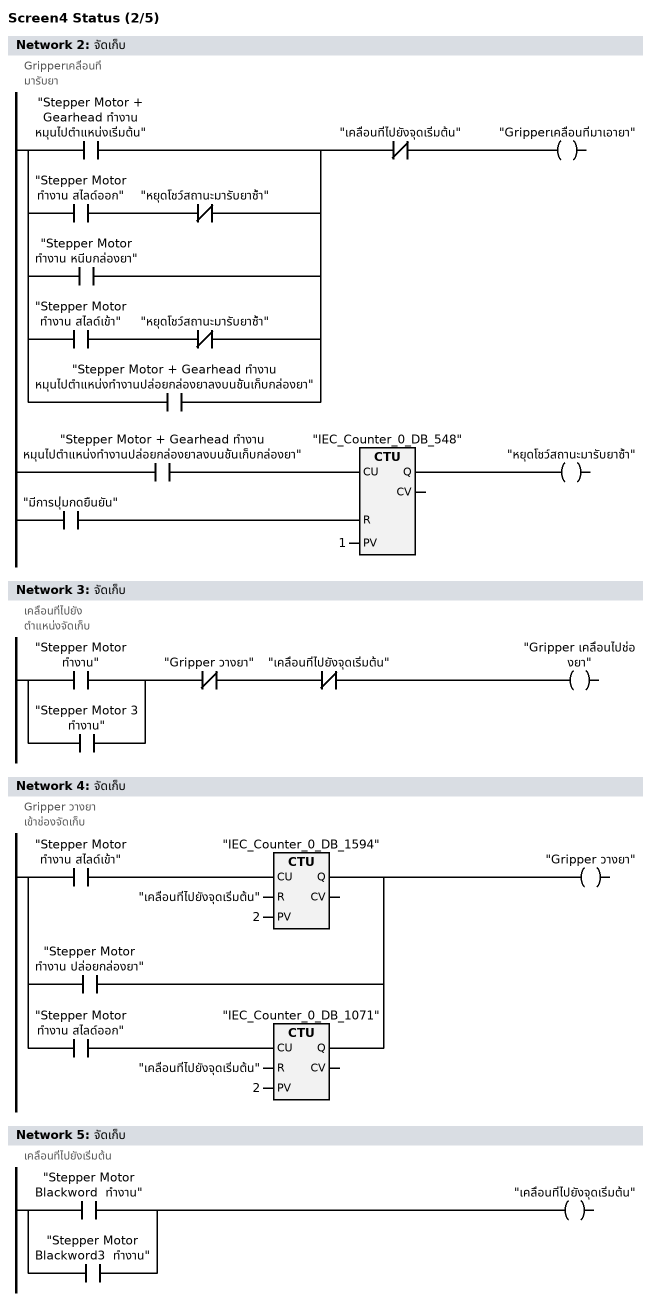
   "Gripperเคลื่อนที่มาเอายา" := ("Stepper Motor + Gearhead ทำงาน หมุนไปตำแหน่งเริ่มต้น" OR ("Stepper Motor ทำงาน สไลด์ออก" AND NOT "หยุดโชว์สถานะมารับยาซ้ำ") OR "Stepper Motor ทำงาน หนีบกล่องยา" OR ("Stepper Motor ทำงาน สไลด์เข้า" AND NOT "หยุดโชว์สถานะมารับยาซ้ำ") OR "Stepper Motor + Gearhead ทำงาน หมุนไปตำแหน่งทำงานปล่อยกล่องยาลงบนชั้นเก็บกล่องยา") AND NOT "เคลื่อนที่ไปยังจุดเริ่มต้น";
   "IEC_Counter_0_DB_548".CTU(CU := "Stepper Motor + Gearhead ทำงาน หมุนไปตำแหน่งทำงานปล่อยกล่องยาลงบนชั้นเก็บกล่องยา",
                           R := "มีการปุ่มกดยืนยัน",
                           PV := 1);
   "หยุดโชว์สถานะมารับยาซ้ำ" := "IEC_Counter_0_DB_548".Q;
END_REGION

REGION Network 3: จัดเก็บ
   // เคลื่อนที่ไปยัง
   // ตำแหน่งจัดเก็บ
   RUNG wire#powerrail
      Contact( "Stepper Motor  ทำงาน" )
      wire#w1
      I_Contact( "Gripper วางยา" )
      I_Contact( "เคลื่อนที่ไปยังจุดเริ่มต้น" )
      Coil( "Gripper เคลื่อนไปช่องยา" )
   END_RUNG
   RUNG wire#powerrail
      Contact( "Stepper Motor 3 ทำงาน" )
   END_RUNG wire#w1
   // the same network as SCL:
   "Gripper เคลื่อนไปช่องยา" := ("Stepper Motor  ทำงาน" OR "Stepper Motor 3 ทำงาน") AND NOT "Gripper วางยา" AND NOT "เคลื่อนที่ไปยังจุดเริ่มต้น";
END_REGION

REGION Network 4: จัดเก็บ
   // Gripper วางยา
   // เข้าช่องจัดเก็บ
   "IEC_Counter_0_DB_1594".CTU(CU := "Stepper Motor ทำงาน สไลด์เข้า",
                           R := "เคลื่อนที่ไปยังจุดเริ่มต้น",
                           PV := 2);
   "IEC_Counter_0_DB_1071".CTU(CU := "Stepper Motor ทำงาน สไลด์ออก", R := "เคลื่อนที่ไปยังจุดเริ่มต้น", PV := 2);
   "Gripper วางยา" := "IEC_Counter_0_DB_1594".Q OR "Stepper Motor ทำงาน ปล่อยกล่องยา" OR "IEC_Counter_0_DB_1071".Q;
END_REGION

REGION Network 5: จัดเก็บ
   // เคลื่อนที่ไปยังเริ่มต้น
   RUNG wire#powerrail
      Contact( "Stepper Motor Blackword  ทำงาน" )
      wire#w1
      Coil( "เคลื่อนที่ไปยังจุดเริ่มต้น" )
   END_RUNG
   RUNG wire#powerrail
      Contact( "Stepper Motor Blackword3  ทำงาน" )
   END_RUNG wire#w1
   // the same network as SCL:
   "เคลื่อนที่ไปยังจุดเริ่มต้น" := "Stepper Motor Blackword  ทำงาน" OR "Stepper Motor Blackword3  ทำงาน";
END_REGION

REGION Network 6: จัดเก็บ
   // รอรับคำสั่งยา
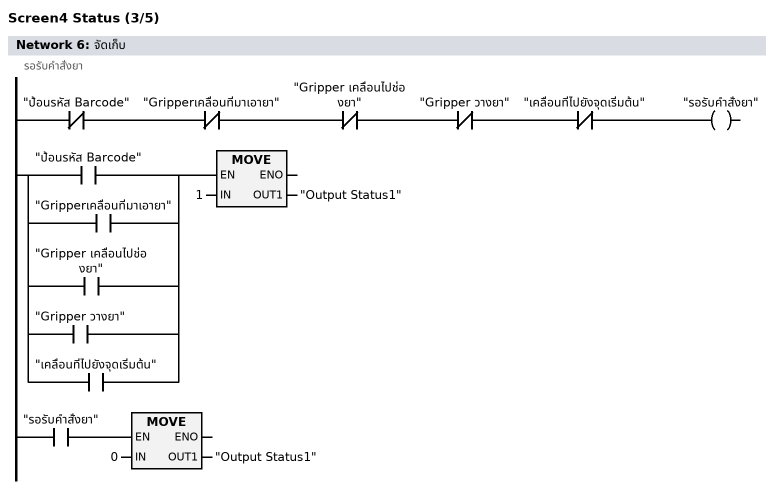
   RUNG wire#powerrail
      I_Contact( "ป้อนรหัส Barcode" )
      I_Contact( "Gripperเคลื่อนที่มาเอายา" )
      I_Contact( "Gripper เคลื่อนไปช่องยา" )
      I_Contact( "Gripper วางยา" )
      I_Contact( "เคลื่อนที่ไปยังจุดเริ่มต้น" )
      Coil( "รอรับคำสั่งยา" )
   END_RUNG
   RUNG wire#powerrail
      Contact( "ป้อนรหัส Barcode" )
      wire#w1
      Move(in := 1, out1 => "Output Status1")
   END_RUNG
   RUNG wire#powerrail
      Contact( "Gripperเคลื่อนที่มาเอายา" )
   END_RUNG wire#w1
   RUNG wire#powerrail
      Contact( "Gripper เคลื่อนไปช่องยา" )
   END_RUNG wire#w1
   RUNG wire#powerrail
      Contact( "Gripper วางยา" )
   END_RUNG wire#w1
   RUNG wire#powerrail
      Contact( "เคลื่อนที่ไปยังจุดเริ่มต้น" )
   END_RUNG wire#w1
   RUNG wire#powerrail
      Contact( "รอรับคำสั่งยา" )
      Move(in := 0, out1 => "Output Status1")
   END_RUNG
   // the same network as SCL:
   "รอรับคำสั่งยา" := NOT "ป้อนรหัส Barcode" AND NOT "Gripperเคลื่อนที่มาเอายา" AND NOT "Gripper เคลื่อนไปช่องยา" AND NOT "Gripper วางยา" AND NOT "เคลื่อนที่ไปยังจุดเริ่มต้น";
   IF "ป้อนรหัส Barcode" OR "Gripperเคลื่อนที่มาเอายา" OR "Gripper เคลื่อนไปช่องยา" OR "Gripper วางยา" OR "เคลื่อนที่ไปยังจุดเริ่มต้น" THEN
       "Output Status1" := 1;
   END_IF;
   IF "รอรับคำสั่งยา" THEN "Output Status1" := 0; END_IF;
END_REGION

REGION Network 7: เบิกจ่าย
   // รับคำสั่งเบิกยา
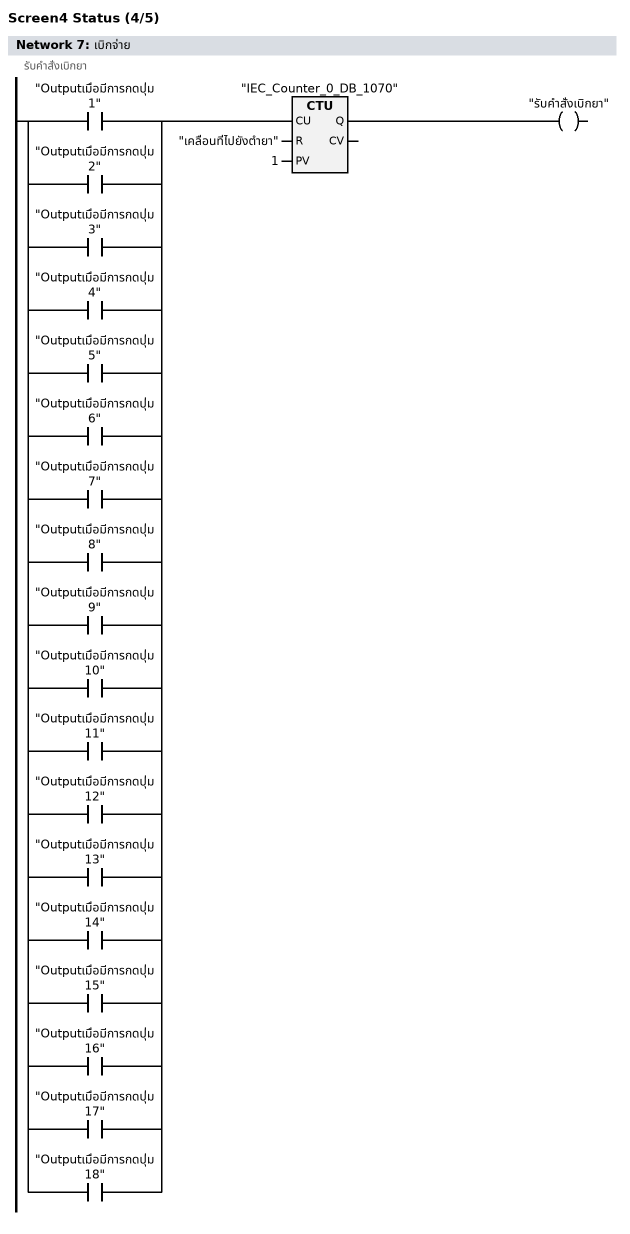
   "IEC_Counter_0_DB_1070".CTU(CU := "Outputเมื่อมีการกดปุ่ม 1" OR "Outputเมื่อมีการกดปุ่ม 2" OR "Outputเมื่อมีการกดปุ่ม 3" OR "Outputเมื่อมีการกดปุ่ม 4" OR "Outputเมื่อมีการกดปุ่ม 5" OR "Outputเมื่อมีการกดปุ่ม 6" OR "Outputเมื่อมีการกดปุ่ม 7" OR "Outputเมื่อมีการกดปุ่ม 8" OR "Outputเมื่อมีการกดปุ่ม 9" OR "Outputเมื่อมีการกดปุ่ม 10" OR "Outputเมื่อมีการกดปุ่ม 11" OR "Outputเมื่อมีการกดปุ่ม 12" OR "Outputเมื่อมีการกดปุ่ม 13" OR "Outputเมื่อมีการกดปุ่ม 14" OR "Outputเมื่อมีการกดปุ่ม 15" OR "Outputเมื่อมีการกดปุ่ม 16" OR "Outputเมื่อมีการกดปุ่ม 17" OR "Outputเมื่อมีการกดปุ่ม 18",
                           R := "เคลื่อนที่ไปยังตำยา",
                           PV := 1);
   "รับคำสั่งเบิกยา" := "IEC_Counter_0_DB_1070".Q;
END_REGION

REGION Network 8: เบิกจ่าย
   // เคลื่อนที่ไปยังตำ
   // แหน่งยา
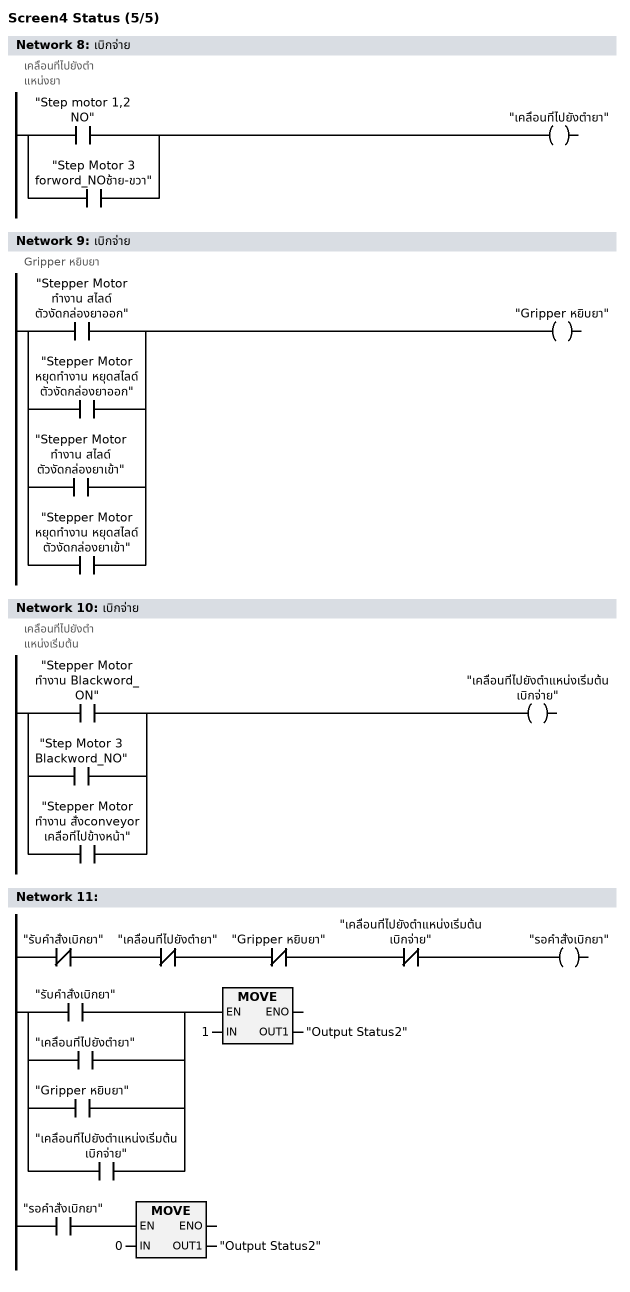
   RUNG wire#powerrail
      Contact( "Step motor 1,2 NO" )
      wire#w1
      Coil( "เคลื่อนที่ไปยังตำยา" )
   END_RUNG
   RUNG wire#powerrail
      Contact( "Step Motor 3 forword_NOซ้าย-ขวา" )
   END_RUNG wire#w1
   // the same network as SCL:
   "เคลื่อนที่ไปยังตำยา" := "Step motor 1,2 NO" OR "Step Motor 3 forword_NOซ้าย-ขวา";
END_REGION

REGION Network 9: เบิกจ่าย
   // Gripper หยิบยา
   RUNG wire#powerrail
      Contact( "Stepper Motor ทำงาน สไลด์ ตัวงัดกล่องยาออก" )
      wire#w1
      Coil( "Gripper หยิบยา" )
   END_RUNG
   RUNG wire#powerrail
      Contact( "Stepper Motor หยุดทำงาน หยุดสไลด์ ตัวงัดกล่องยาออก" )
   END_RUNG wire#w1
   RUNG wire#powerrail
      Contact( "Stepper Motor ทำงาน สไลด์ ตัวงัดกล่องยาเข้า" )
   END_RUNG wire#w1
   RUNG wire#powerrail
      Contact( "Stepper Motor หยุดทำงาน หยุดสไลด์ ตัวงัดกล่องยาเข้า" )
   END_RUNG wire#w1
   // the same network as SCL:
   "Gripper หยิบยา" := "Stepper Motor ทำงาน สไลด์ ตัวงัดกล่องยาออก" OR "Stepper Motor หยุดทำงาน หยุดสไลด์ ตัวงัดกล่องยาออก" OR "Stepper Motor ทำงาน สไลด์ ตัวงัดกล่องยาเข้า" OR "Stepper Motor หยุดทำงาน หยุดสไลด์ ตัวงัดกล่องยาเข้า";
END_REGION

REGION Network 10: เบิกจ่าย
   // เคลื่อนที่ไปยังตำ
   // แหน่งเริ่มต้น
   RUNG wire#powerrail
      Contact( "Stepper Motor  ทำงาน Blackword_ON" )
      wire#w1
      Coil( "เคลื่อนที่ไปยังตำแหน่งเริ่มต้น เบิกจ่าย" )
   END_RUNG
   RUNG wire#powerrail
      Contact( "Step Motor 3 Blackword_NO" )
   END_RUNG wire#w1
   RUNG wire#powerrail
      Contact( "Stepper Motor ทำงาน สั่งconveyor เคลื่อที่ไปข้างหน้า" )
   END_RUNG wire#w1
   // the same network as SCL:
   "เคลื่อนที่ไปยังตำแหน่งเริ่มต้น เบิกจ่าย" := "Stepper Motor  ทำงาน Blackword_ON" OR "Step Motor 3 Blackword_NO" OR "Stepper Motor ทำงาน สั่งconveyor เคลื่อที่ไปข้างหน้า";
END_REGION

REGION Network 11
   RUNG wire#powerrail
      I_Contact( "รับคำสั่งเบิกยา" )
      I_Contact( "เคลื่อนที่ไปยังตำยา" )
      I_Contact( "Gripper หยิบยา" )
      I_Contact( "เคลื่อนที่ไปยังตำแหน่งเริ่มต้น เบิกจ่าย" )
      Coil( "รอคำสั่งเบิกยา" )
   END_RUNG
   RUNG wire#powerrail
      Contact( "รับคำสั่งเบิกยา" )
      wire#w1
      Move(in := 1, out1 => "Output Status2")
   END_RUNG
   RUNG wire#powerrail
      Contact( "เคลื่อนที่ไปยังตำยา" )
   END_RUNG wire#w1
   RUNG wire#powerrail
      Contact( "Gripper หยิบยา" )
   END_RUNG wire#w1
   RUNG wire#powerrail
      Contact( "เคลื่อนที่ไปยังตำแหน่งเริ่มต้น เบิกจ่าย" )
   END_RUNG wire#w1
   RUNG wire#powerrail
      Contact( "รอคำสั่งเบิกยา" )
      Move(in := 0, out1 => "Output Status2")
   END_RUNG
   // the same network as SCL:
   "รอคำสั่งเบิกยา" := NOT "รับคำสั่งเบิกยา" AND NOT "เคลื่อนที่ไปยังตำยา" AND NOT "Gripper หยิบยา" AND NOT "เคลื่อนที่ไปยังตำแหน่งเริ่มต้น เบิกจ่าย";
   IF "รับคำสั่งเบิกยา" OR "เคลื่อนที่ไปยังตำยา" OR "Gripper หยิบยา" OR "เคลื่อนที่ไปยังตำแหน่งเริ่มต้น เบิกจ่าย" THEN
       "Output Status2" := 1;
   END_IF;
   IF "รอคำสั่งเบิกยา" THEN "Output Status2" := 0; END_IF;
END_REGION
END_FUNCTION

// folder: Screen หน้าจอ/Conveyor

FUNCTION "Conveyor" : Void   // FC1, LAD
{ S7_Optimized_Access := 'TRUE' }
VERSION : 0.1
   VAR_INPUT
      "เวลาที่Brushless Motor ทำงาน" : Time;
   END_VAR
   VAR_OUTPUT
      "OutputหลังPhotoelectic sensor 3 ตรวจเจอวัตถุ" : Bool;
   END_VAR
BEGIN

REGION Network 1
